// --- Siemens Structured Format ---
DATA_BLOCK "model__HS32_IW50_"
{ S7_Optimized_Access := 'TRUE' }
VERSION :
NON_RETAIN
   VAR
      W_i : ARRAY[0..31, 0..39] OF REAL;
      W_f : ARRAY[0..31, 0..39] OF REAL;
      W_g : ARRAY[0..31, 0..39] OF REAL;
      W_o : ARRAY[0..31, 0..39] OF REAL;
      R_i : ARRAY[0..31, 0..31] OF REAL;
      R_f : ARRAY[0..31, 0..31] OF REAL;
      R_g : ARRAY[0..31, 0..31] OF REAL;
      R_o : ARRAY[0..31, 0..31] OF REAL;
      B_i : ARRAY[0..31] OF REAL;
      B_f : ARRAY[0..31] OF REAL;
      B_g : ARRAY[0..31] OF REAL;
      B_o : ARRAY[0..31] OF REAL;
      FC_W : ARRAY[0..39, 0..31] OF REAL;
      FC_B : ARRAY[0..39] OF REAL;
   END_VAR
BEGIN

      W_i[0,0] := 0.03335211;
      W_i[0,1] := 0.01294965;
      W_i[0,2] := -0.02368959;
      W_i[0,3] := 0.02531582;
      W_i[0,4] := -0.09620859;
      W_i[0,5] := -0.01378066;
      W_i[0,6] := 0.03223424;
      W_i[0,7] := 0.44872370;
      W_i[0,8] := 0.10217454;
      W_i[0,9] := -0.36218736;
      W_i[0,10] := 0.04811719;
      W_i[0,11] := -0.30795375;
      W_i[0,12] := -0.13306537;
      W_i[0,13] := -0.13929474;
      W_i[0,14] := -0.02903975;
      W_i[0,15] := 0.11072005;
      W_i[0,16] := 0.03733860;
      W_i[0,17] := 0.00262149;
      W_i[0,18] := 0.23541802;
      W_i[0,19] := 0.20732951;
      W_i[0,20] := 0.04801108;
      W_i[0,21] := -0.28304836;
      W_i[0,22] := -0.50957590;
      W_i[0,23] := 0.04589643;
      W_i[0,24] := -0.43349111;
      W_i[0,25] := -0.42231610;
      W_i[0,26] := 0.15247093;
      W_i[0,27] := 0.29900289;
      W_i[0,28] := 0.08071815;
      W_i[0,29] := 0.16624704;
      W_i[0,30] := -0.21118966;
      W_i[0,31] := -0.06602232;
      W_i[0,32] := 0.02604864;
      W_i[0,33] := -0.14019786;
      W_i[0,34] := -0.40027091;
      W_i[0,35] := 0.18787135;
      W_i[0,36] := 0.02354476;
      W_i[0,37] := 0.16503902;
      W_i[0,38] := -0.08474749;
      W_i[0,39] := 0.36904612;
      W_i[1,0] := -0.04397624;
      W_i[1,1] := 0.12521634;
      W_i[1,2] := 0.00926329;
      W_i[1,3] := 0.07923686;
      W_i[1,4] := -0.48040998;
      W_i[1,5] := 0.11951946;
      W_i[1,6] := -0.05899520;
      W_i[1,7] := 0.08414336;
      W_i[1,8] := -0.05504049;
      W_i[1,9] := -0.01812936;
      W_i[1,10] := -0.07156652;
      W_i[1,11] := -0.13873386;
      W_i[1,12] := -0.06473546;
      W_i[1,13] := -0.01150122;
      W_i[1,14] := 0.01369441;
      W_i[1,15] := -0.04945480;
      W_i[1,16] := 0.03672740;
      W_i[1,17] := -0.01182620;
      W_i[1,18] := 0.05847014;
      W_i[1,19] := 0.12310074;
      W_i[1,20] := 0.00140591;
      W_i[1,21] := 0.05102165;
      W_i[1,22] := 0.02194597;
      W_i[1,23] := 0.02794340;
      W_i[1,24] := -0.11971385;
      W_i[1,25] := 0.01236170;
      W_i[1,26] := 0.02725715;
      W_i[1,27] := -0.16358410;
      W_i[1,28] := 0.09302291;
      W_i[1,29] := -0.07609808;
      W_i[1,30] := 0.12344577;
      W_i[1,31] := 0.27449563;
      W_i[1,32] := 0.19618334;
      W_i[1,33] := -0.13863903;
      W_i[1,34] := -0.14182809;
      W_i[1,35] := -0.04518571;
      W_i[1,36] := -0.11997688;
      W_i[1,37] := 0.13018343;
      W_i[1,38] := 0.03084990;
      W_i[1,39] := 0.01552542;
      W_i[2,0] := -0.06228839;
      W_i[2,1] := 0.31358635;
      W_i[2,2] := -0.02805484;
      W_i[2,3] := 0.06225382;
      W_i[2,4] := -0.10929245;
      W_i[2,5] := 0.09066710;
      W_i[2,6] := -0.09841387;
      W_i[2,7] := 0.21516874;
      W_i[2,8] := -0.04192384;
      W_i[2,9] := -0.24015123;
      W_i[2,10] := 0.18081841;
      W_i[2,11] := -0.22261326;
      W_i[2,12] := 0.15341285;
      W_i[2,13] := -0.01613901;
      W_i[2,14] := 0.00278526;
      W_i[2,15] := 0.00110682;
      W_i[2,16] := 0.01401542;
      W_i[2,17] := 0.00157240;
      W_i[2,18] := -0.00937896;
      W_i[2,19] := 0.08156285;
      W_i[2,20] := -0.10387972;
      W_i[2,21] := 0.07669238;
      W_i[2,22] := 0.10504947;
      W_i[2,23] := 0.02962043;
      W_i[2,24] := 0.06015503;
      W_i[2,25] := -0.38022354;
      W_i[2,26] := 0.01376416;
      W_i[2,27] := -0.19910932;
      W_i[2,28] := -0.11147632;
      W_i[2,29] := -0.06024737;
      W_i[2,30] := 0.33740976;
      W_i[2,31] := -0.14441007;
      W_i[2,32] := 0.09709183;
      W_i[2,33] := -0.01737254;
      W_i[2,34] := 0.10466792;
      W_i[2,35] := -0.13491732;
      W_i[2,36] := 0.03209321;
      W_i[2,37] := -0.20953350;
      W_i[2,38] := 0.02072377;
      W_i[2,39] := -0.03477554;
      W_i[3,0] := -0.20035338;
      W_i[3,1] := -0.05025988;
      W_i[3,2] := -0.08164182;
      W_i[3,3] := -0.08261910;
      W_i[3,4] := 0.24175876;
      W_i[3,5] := -0.19314556;
      W_i[3,6] := 0.16183864;
      W_i[3,7] := -0.53965092;
      W_i[3,8] := 0.12166216;
      W_i[3,9] := 0.06300285;
      W_i[3,10] := 0.24695574;
      W_i[3,11] := -0.06766498;
      W_i[3,12] := -0.10851647;
      W_i[3,13] := -0.09679550;
      W_i[3,14] := 0.19846407;
      W_i[3,15] := 0.24224226;
      W_i[3,16] := -0.04479418;
      W_i[3,17] := 0.09416196;
      W_i[3,18] := -0.05448310;
      W_i[3,19] := -0.14848493;
      W_i[3,20] := -0.13104467;
      W_i[3,21] := 0.01169914;
      W_i[3,22] := 0.13594244;
      W_i[3,23] := -0.09969987;
      W_i[3,24] := -0.51131010;
      W_i[3,25] := -0.49498364;
      W_i[3,26] := -0.00815858;
      W_i[3,27] := -0.01644909;
      W_i[3,28] := -0.31252897;
      W_i[3,29] := -0.13085435;
      W_i[3,30] := 0.42893934;
      W_i[3,31] := -0.31215337;
      W_i[3,32] := -0.04756459;
      W_i[3,33] := -0.18021715;
      W_i[3,34] := -0.17681709;
      W_i[3,35] := -0.15721944;
      W_i[3,36] := 0.22830988;
      W_i[3,37] := 0.15386219;
      W_i[3,38] := -0.11364616;
      W_i[3,39] := 0.85980165;
      W_i[4,0] := -0.05922852;
      W_i[4,1] := 0.47120315;
      W_i[4,2] := 0.31002536;
      W_i[4,3] := 0.05706808;
      W_i[4,4] := 0.21668130;
      W_i[4,5] := 0.09678623;
      W_i[4,6] := 0.37920210;
      W_i[4,7] := 0.11913582;
      W_i[4,8] := 0.18588071;
      W_i[4,9] := -0.54219109;
      W_i[4,10] := 0.27432936;
      W_i[4,11] := -0.28996110;
      W_i[4,12] := 0.63514346;
      W_i[4,13] := 0.18675460;
      W_i[4,14] := 0.04656186;
      W_i[4,15] := 0.13881819;
      W_i[4,16] := -0.17344026;
      W_i[4,17] := 0.07573078;
      W_i[4,18] := 0.08432268;
      W_i[4,19] := -0.39324254;
      W_i[4,20] := 0.22332989;
      W_i[4,21] := 0.55870950;
      W_i[4,22] := -0.48373845;
      W_i[4,23] := -0.31563666;
      W_i[4,24] := 0.31388757;
      W_i[4,25] := 0.28351381;
      W_i[4,26] := 0.00493392;
      W_i[4,27] := -0.14279558;
      W_i[4,28] := 0.01328408;
      W_i[4,29] := -0.13343237;
      W_i[4,30] := -0.52480948;
      W_i[4,31] := -0.44383386;
      W_i[4,32] := -0.22764747;
      W_i[4,33] := 0.36674559;
      W_i[4,34] := 0.28135881;
      W_i[4,35] := -0.37915036;
      W_i[4,36] := 0.29197508;
      W_i[4,37] := -0.36793157;
      W_i[4,38] := 0.61301214;
      W_i[4,39] := 0.29268816;
      W_i[5,0] := -0.15593423;
      W_i[5,1] := -0.08324785;
      W_i[5,2] := 0.00935801;
      W_i[5,3] := 0.08572404;
      W_i[5,4] := -0.04179911;
      W_i[5,5] := -0.08974203;
      W_i[5,6] := -0.03267067;
      W_i[5,7] := -0.12864745;
      W_i[5,8] := 0.03684423;
      W_i[5,9] := -0.13796446;
      W_i[5,10] := 0.05928193;
      W_i[5,11] := -0.19078448;
      W_i[5,12] := 0.04955722;
      W_i[5,13] := -0.13951716;
      W_i[5,14] := 0.01461054;
      W_i[5,15] := 0.05807864;
      W_i[5,16] := -0.02155071;
      W_i[5,17] := 0.06774671;
      W_i[5,18] := -0.00056143;
      W_i[5,19] := 0.02993268;
      W_i[5,20] := -0.04689442;
      W_i[5,21] := 0.14087728;
      W_i[5,22] := -0.00434205;
      W_i[5,23] := -0.14380206;
      W_i[5,24] := -0.53344935;
      W_i[5,25] := 0.06604308;
      W_i[5,26] := 0.23374112;
      W_i[5,27] := 0.02832700;
      W_i[5,28] := 0.09275237;
      W_i[5,29] := 0.07908134;
      W_i[5,30] := -0.10972932;
      W_i[5,31] := -0.08337840;
      W_i[5,32] := 0.04662216;
      W_i[5,33] := -0.03259875;
      W_i[5,34] := 0.17782964;
      W_i[5,35] := 0.18201338;
      W_i[5,36] := 0.00404544;
      W_i[5,37] := 0.04663613;
      W_i[5,38] := 0.13219389;
      W_i[5,39] := -0.00446346;
      W_i[6,0] := 0.10576568;
      W_i[6,1] := 0.05325136;
      W_i[6,2] := -0.05492130;
      W_i[6,3] := -0.11396622;
      W_i[6,4] := 0.02959487;
      W_i[6,5] := 0.04510606;
      W_i[6,6] := 0.21042347;
      W_i[6,7] := 0.11686674;
      W_i[6,8] := 0.17569162;
      W_i[6,9] := -0.22145574;
      W_i[6,10] := 0.01603481;
      W_i[6,11] := -0.21858092;
      W_i[6,12] := 0.03767690;
      W_i[6,13] := -0.15889299;
      W_i[6,14] := 0.02401877;
      W_i[6,15] := -0.09354293;
      W_i[6,16] := -0.06953581;
      W_i[6,17] := 0.01671052;
      W_i[6,18] := 0.14821531;
      W_i[6,19] := 0.03779463;
      W_i[6,20] := 0.31719235;
      W_i[6,21] := 0.26848948;
      W_i[6,22] := 0.24316274;
      W_i[6,23] := -0.03367342;
      W_i[6,24] := -0.43727583;
      W_i[6,25] := -0.31479907;
      W_i[6,26] := 0.40017867;
      W_i[6,27] := -0.00208360;
      W_i[6,28] := 0.18425919;
      W_i[6,29] := 0.37186173;
      W_i[6,30] := 0.17230935;
      W_i[6,31] := -0.07113405;
      W_i[6,32] := 0.06234986;
      W_i[6,33] := -0.04395010;
      W_i[6,34] := 0.03162268;
      W_i[6,35] := 0.12794030;
      W_i[6,36] := -0.06928633;
      W_i[6,37] := 0.28019226;
      W_i[6,38] := -0.08624983;
      W_i[6,39] := -0.05943641;
      W_i[7,0] := 0.24273345;
      W_i[7,1] := 0.02628726;
      W_i[7,2] := -0.37892520;
      W_i[7,3] := 0.15462431;
      W_i[7,4] := -0.06835640;
      W_i[7,5] := -0.01244921;
      W_i[7,6] := -0.13799721;
      W_i[7,7] := 0.00364937;
      W_i[7,8] := -0.11085126;
      W_i[7,9] := -0.08217847;
      W_i[7,10] := 0.06155964;
      W_i[7,11] := 0.00664949;
      W_i[7,12] := -0.21111001;
      W_i[7,13] := -0.09906641;
      W_i[7,14] := 0.01441233;
      W_i[7,15] := 0.05717637;
      W_i[7,16] := -0.01254125;
      W_i[7,17] := -0.00084031;
      W_i[7,18] := 0.75006574;
      W_i[7,19] := 0.04177287;
      W_i[7,20] := -0.16489621;
      W_i[7,21] := -0.11358984;
      W_i[7,22] := -0.32568359;
      W_i[7,23] := -0.05461695;
      W_i[7,24] := -0.68117988;
      W_i[7,25] := -0.38877121;
      W_i[7,26] := 0.21966200;
      W_i[7,27] := 0.08412468;
      W_i[7,28] := -0.18800470;
      W_i[7,29] := -0.37555104;
      W_i[7,30] := -0.20995075;
      W_i[7,31] := -0.00920301;
      W_i[7,32] := -0.38933340;
      W_i[7,33] := 0.03684454;
      W_i[7,34] := -0.00580212;
      W_i[7,35] := -0.12717755;
      W_i[7,36] := 0.00740355;
      W_i[7,37] := -0.09031770;
      W_i[7,38] := -0.11013316;
      W_i[7,39] := -0.04330545;
      W_i[8,0] := -0.06802954;
      W_i[8,1] := -0.02636882;
      W_i[8,2] := 0.04332832;
      W_i[8,3] := -0.12407507;
      W_i[8,4] := 0.01348176;
      W_i[8,5] := -0.07925858;
      W_i[8,6] := -0.00761013;
      W_i[8,7] := 0.03581184;
      W_i[8,8] := 0.02980794;
      W_i[8,9] := -0.13043974;
      W_i[8,10] := 0.09170759;
      W_i[8,11] := -0.16562377;
      W_i[8,12] := -0.12424939;
      W_i[8,13] := 0.05662967;
      W_i[8,14] := -0.21820237;
      W_i[8,15] := 0.03667807;
      W_i[8,16] := 0.01659469;
      W_i[8,17] := 0.00193780;
      W_i[8,18] := -0.03699196;
      W_i[8,19] := -0.02531029;
      W_i[8,20] := -0.00570031;
      W_i[8,21] := 0.10410964;
      W_i[8,22] := 0.06439263;
      W_i[8,23] := -0.07894669;
      W_i[8,24] := -0.28273982;
      W_i[8,25] := -0.23450002;
      W_i[8,26] := 0.05201263;
      W_i[8,27] := -0.03252214;
      W_i[8,28] := -0.01173223;
      W_i[8,29] := 0.14622457;
      W_i[8,30] := 0.17911775;
      W_i[8,31] := -0.11378439;
      W_i[8,32] := 0.07194026;
      W_i[8,33] := 0.01723621;
      W_i[8,34] := 0.30313444;
      W_i[8,35] := 0.11768141;
      W_i[8,36] := -0.01293503;
      W_i[8,37] := -0.00394995;
      W_i[8,38] := -0.14124557;
      W_i[8,39] := 0.13445212;
      W_i[9,0] := 0.41246179;
      W_i[9,1] := -0.12685674;
      W_i[9,2] := -0.45634085;
      W_i[9,3] := -0.20486909;
      W_i[9,4] := -0.07218436;
      W_i[9,5] := -0.09485383;
      W_i[9,6] := 0.19853495;
      W_i[9,7] := 0.07240235;
      W_i[9,8] := -0.04039089;
      W_i[9,9] := -0.09886632;
      W_i[9,10] := -0.11097286;
      W_i[9,11] := -0.28303620;
      W_i[9,12] := 0.15636595;
      W_i[9,13] := 0.12219298;
      W_i[9,14] := 0.16322424;
      W_i[9,15] := 0.06697550;
      W_i[9,16] := -0.11505034;
      W_i[9,17] := 0.01392226;
      W_i[9,18] := -0.03821991;
      W_i[9,19] := 0.35102692;
      W_i[9,20] := 0.15118374;
      W_i[9,21] := 0.24640937;
      W_i[9,22] := 0.02153728;
      W_i[9,23] := -0.02444457;
      W_i[9,24] := 0.13131861;
      W_i[9,25] := -0.16178758;
      W_i[9,26] := -0.05835283;
      W_i[9,27] := -0.28876659;
      W_i[9,28] := -0.22485775;
      W_i[9,29] := -0.10750232;
      W_i[9,30] := 0.07209923;
      W_i[9,31] := -0.16665789;
      W_i[9,32] := 0.09024238;
      W_i[9,33] := 0.15630057;
      W_i[9,34] := 0.22654596;
      W_i[9,35] := -0.16981296;
      W_i[9,36] := 0.09843912;
      W_i[9,37] := -0.08633557;
      W_i[9,38] := 0.06714951;
      W_i[9,39] := -0.10012744;
      W_i[10,0] := 0.06098233;
      W_i[10,1] := 0.00406449;
      W_i[10,2] := -0.07085112;
      W_i[10,3] := -0.38051835;
      W_i[10,4] := -0.14092854;
      W_i[10,5] := -0.05471934;
      W_i[10,6] := -0.09075350;
      W_i[10,7] := 0.09081808;
      W_i[10,8] := 0.07290499;
      W_i[10,9] := 0.21984702;
      W_i[10,10] := -0.00319992;
      W_i[10,11] := -0.87133026;
      W_i[10,12] := 0.25286415;
      W_i[10,13] := -0.20190343;
      W_i[10,14] := -0.29993787;
      W_i[10,15] := -0.01450086;
      W_i[10,16] := -0.04255661;
      W_i[10,17] := 0.50596321;
      W_i[10,18] := -0.03224555;
      W_i[10,19] := 0.00962685;
      W_i[10,20] := 0.02170906;
      W_i[10,21] := 0.00463841;
      W_i[10,22] := 0.00428250;
      W_i[10,23] := 0.02700867;
      W_i[10,24] := -0.49260652;
      W_i[10,25] := -0.60828519;
      W_i[10,26] := 0.08981935;
      W_i[10,27] := -0.05126838;
      W_i[10,28] := 0.10806957;
      W_i[10,29] := 0.06330517;
      W_i[10,30] := 0.09711373;
      W_i[10,31] := -0.19667481;
      W_i[10,32] := 0.04281054;
      W_i[10,33] := 0.06612559;
      W_i[10,34] := -0.12514877;
      W_i[10,35] := 0.09477433;
      W_i[10,36] := 0.02109047;
      W_i[10,37] := 0.06420635;
      W_i[10,38] := 0.06682578;
      W_i[10,39] := 0.70137119;
      W_i[11,0] := -0.19831482;
      W_i[11,1] := -0.10508762;
      W_i[11,2] := 0.14985219;
      W_i[11,3] := -0.25513422;
      W_i[11,4] := 0.22445941;
      W_i[11,5] := -0.17102213;
      W_i[11,6] := 0.03812301;
      W_i[11,7] := 0.06178447;
      W_i[11,8] := -0.06147041;
      W_i[11,9] := 0.01455363;
      W_i[11,10] := 0.21236670;
      W_i[11,11] := -0.06561671;
      W_i[11,12] := -0.23426783;
      W_i[11,13] := 0.09121598;
      W_i[11,14] := -0.11325682;
      W_i[11,15] := 0.14043726;
      W_i[11,16] := -0.03869899;
      W_i[11,17] := 0.07733488;
      W_i[11,18] := -0.00199524;
      W_i[11,19] := 0.05081591;
      W_i[11,20] := -0.45575571;
      W_i[11,21] := -0.48401207;
      W_i[11,22] := -0.20732693;
      W_i[11,23] := -0.15296169;
      W_i[11,24] := -0.30430803;
      W_i[11,25] := -0.48835382;
      W_i[11,26] := -0.19211042;
      W_i[11,27] := 0.21992902;
      W_i[11,28] := -0.36160839;
      W_i[11,29] := -0.36730286;
      W_i[11,30] := -0.27825427;
      W_i[11,31] := 0.49533325;
      W_i[11,32] := 0.01973951;
      W_i[11,33] := 0.13294254;
      W_i[11,34] := -0.31377479;
      W_i[11,35] := 0.01389581;
      W_i[11,36] := -0.10732657;
      W_i[11,37] := -0.10178760;
      W_i[11,38] := -0.04468285;
      W_i[11,39] := 0.88543254;
      W_i[12,0] := -0.07785182;
      W_i[12,1] := -0.02275736;
      W_i[12,2] := -0.01598639;
      W_i[12,3] := -0.28018406;
      W_i[12,4] := 0.04472728;
      W_i[12,5] := -0.07362497;
      W_i[12,6] := 0.10421625;
      W_i[12,7] := 0.29120883;
      W_i[12,8] := 0.07516699;
      W_i[12,9] := -0.19484363;
      W_i[12,10] := 0.04389035;
      W_i[12,11] := 0.07964118;
      W_i[12,12] := 0.04882551;
      W_i[12,13] := -0.09314007;
      W_i[12,14] := -0.00104783;
      W_i[12,15] := 0.12430931;
      W_i[12,16] := -0.00889617;
      W_i[12,17] := -0.00109596;
      W_i[12,18] := 0.93196803;
      W_i[12,19] := 0.07360591;
      W_i[12,20] := -0.04771593;
      W_i[12,21] := 0.00891263;
      W_i[12,22] := -0.22154218;
      W_i[12,23] := -0.00681991;
      W_i[12,24] := -0.28159559;
      W_i[12,25] := -0.33888876;
      W_i[12,26] := 0.11433282;
      W_i[12,27] := -0.10486361;
      W_i[12,28] := -0.09925523;
      W_i[12,29] := -0.00571722;
      W_i[12,30] := -0.36633971;
      W_i[12,31] := -0.06006427;
      W_i[12,32] := -0.22424956;
      W_i[12,33] := -0.32570857;
      W_i[12,34] := -0.57398140;
      W_i[12,35] := 0.05099113;
      W_i[12,36] := 0.00469301;
      W_i[12,37] := 0.02404906;
      W_i[12,38] := 0.01321469;
      W_i[12,39] := -0.01789427;
      W_i[13,0] := 0.13228506;
      W_i[13,1] := 0.10746437;
      W_i[13,2] := -0.02473475;
      W_i[13,3] := -0.01283106;
      W_i[13,4] := -0.11313344;
      W_i[13,5] := 0.01196120;
      W_i[13,6] := -0.10874924;
      W_i[13,7] := -0.09509301;
      W_i[13,8] := 0.00865637;
      W_i[13,9] := -0.15097018;
      W_i[13,10] := 0.07857790;
      W_i[13,11] := -0.13828419;
      W_i[13,12] := 0.18908830;
      W_i[13,13] := -0.03993330;
      W_i[13,14] := 0.01041046;
      W_i[13,15] := 0.00195818;
      W_i[13,16] := -0.02810182;
      W_i[13,17] := -0.00908193;
      W_i[13,18] := -0.01383985;
      W_i[13,19] := 0.01692491;
      W_i[13,20] := 0.26870248;
      W_i[13,21] := 0.50765073;
      W_i[13,22] := 0.34594440;
      W_i[13,23] := -0.03796029;
      W_i[13,24] := -0.65532976;
      W_i[13,25] := -0.80482006;
      W_i[13,26] := 0.01045384;
      W_i[13,27] := -0.46558616;
      W_i[13,28] := 0.19693999;
      W_i[13,29] := 0.14626113;
      W_i[13,30] := 0.43212712;
      W_i[13,31] := 0.01994485;
      W_i[13,32] := -0.32835758;
      W_i[13,33] := -0.17723863;
      W_i[13,34] := 0.20528001;
      W_i[13,35] := -0.34655216;
      W_i[13,36] := -0.06347063;
      W_i[13,37] := -0.07853378;
      W_i[13,38] := 0.15984800;
      W_i[13,39] := 0.00452000;
      W_i[14,0] := -0.00785071;
      W_i[14,1] := -0.08457682;
      W_i[14,2] := -0.03021882;
      W_i[14,3] := 0.06919254;
      W_i[14,4] := -0.07102513;
      W_i[14,5] := -0.11649032;
      W_i[14,6] := -0.13716960;
      W_i[14,7] := 0.12219854;
      W_i[14,8] := -0.03531046;
      W_i[14,9] := -0.07139499;
      W_i[14,10] := -0.28596520;
      W_i[14,11] := -0.20866406;
      W_i[14,12] := -0.09834762;
      W_i[14,13] := -0.17434466;
      W_i[14,14] := 0.05277216;
      W_i[14,15] := 0.05034710;
      W_i[14,16] := -0.04395842;
      W_i[14,17] := 0.01994520;
      W_i[14,18] := -0.00284745;
      W_i[14,19] := -0.01580888;
      W_i[14,20] := 0.35238999;
      W_i[14,21] := -0.30224216;
      W_i[14,22] := -0.01767650;
      W_i[14,23] := 0.06807997;
      W_i[14,24] := -0.02559922;
      W_i[14,25] := -0.02666317;
      W_i[14,26] := 0.03206453;
      W_i[14,27] := 0.41885376;
      W_i[14,28] := 0.04192250;
      W_i[14,29] := -0.05693231;
      W_i[14,30] := 0.07898923;
      W_i[14,31] := 0.18591896;
      W_i[14,32] := -0.06221836;
      W_i[14,33] := 0.24379699;
      W_i[14,34] := -0.13005574;
      W_i[14,35] := 0.04800267;
      W_i[14,36] := 0.09943730;
      W_i[14,37] := -0.03374345;
      W_i[14,38] := -0.03513518;
      W_i[14,39] := -0.07157569;
      W_i[15,0] := -0.15272453;
      W_i[15,1] := 0.13645852;
      W_i[15,2] := 0.04745365;
      W_i[15,3] := -0.20139949;
      W_i[15,4] := 0.03436549;
      W_i[15,5] := 0.06549827;
      W_i[15,6] := -0.17606948;
      W_i[15,7] := 0.05636362;
      W_i[15,8] := 0.15209863;
      W_i[15,9] := -0.04455522;
      W_i[15,10] := 0.01616382;
      W_i[15,11] := 0.02472791;
      W_i[15,12] := 0.01587282;
      W_i[15,13] := 0.06205805;
      W_i[15,14] := -0.01110538;
      W_i[15,15] := -0.05222612;
      W_i[15,16] := -0.00958592;
      W_i[15,17] := 0.05923622;
      W_i[15,18] := 0.03878036;
      W_i[15,19] := -0.04121817;
      W_i[15,20] := -0.04009682;
      W_i[15,21] := 0.02127116;
      W_i[15,22] := -0.04295387;
      W_i[15,23] := -0.08172908;
      W_i[15,24] := -0.48291191;
      W_i[15,25] := -0.58466184;
      W_i[15,26] := -0.04407280;
      W_i[15,27] := 0.00633614;
      W_i[15,28] := -0.10225561;
      W_i[15,29] := 0.48959246;
      W_i[15,30] := -0.22612220;
      W_i[15,31] := -0.01089828;
      W_i[15,32] := -0.25822705;
      W_i[15,33] := -0.17706192;
      W_i[15,34] := -0.61160076;
      W_i[15,35] := 0.09040477;
      W_i[15,36] := 0.02512925;
      W_i[15,37] := -0.06701392;
      W_i[15,38] := -0.08561996;
      W_i[15,39] := 0.53837699;
      W_i[16,0] := -0.07811758;
      W_i[16,1] := 0.05202470;
      W_i[16,2] := 0.03025672;
      W_i[16,3] := 0.04235693;
      W_i[16,4] := -0.06725603;
      W_i[16,5] := -0.00081394;
      W_i[16,6] := -0.09191743;
      W_i[16,7] := 0.24823768;
      W_i[16,8] := 0.02800119;
      W_i[16,9] := -0.27142274;
      W_i[16,10] := -0.06025495;
      W_i[16,11] := -0.51023978;
      W_i[16,12] := 0.54432988;
      W_i[16,13] := -0.07693134;
      W_i[16,14] := 0.03643584;
      W_i[16,15] := 0.04252481;
      W_i[16,16] := -0.00319035;
      W_i[16,17] := -0.16166179;
      W_i[16,18] := -0.10264453;
      W_i[16,19] := -0.72658694;
      W_i[16,20] := -0.08637008;
      W_i[16,21] := -0.15963581;
      W_i[16,22] := -0.16920443;
      W_i[16,23] := -0.03855850;
      W_i[16,24] := -0.09449768;
      W_i[16,25] := -0.15130939;
      W_i[16,26] := -0.07037468;
      W_i[16,27] := 0.05760185;
      W_i[16,28] := 0.01705931;
      W_i[16,29] := 0.05011314;
      W_i[16,30] := -0.01099099;
      W_i[16,31] := -0.06498095;
      W_i[16,32] := 0.15388052;
      W_i[16,33] := -0.03008743;
      W_i[16,34] := -0.91294670;
      W_i[16,35] := 0.04827264;
      W_i[16,36] := 0.00881240;
      W_i[16,37] := 0.02179604;
      W_i[16,38] := 0.47361013;
      W_i[16,39] := 0.58336878;
      W_i[17,0] := -0.22612889;
      W_i[17,1] := -0.03230098;
      W_i[17,2] := 0.24163076;
      W_i[17,3] := 0.20527579;
      W_i[17,4] := -0.44036463;
      W_i[17,5] := 0.28084049;
      W_i[17,6] := -0.51067066;
      W_i[17,7] := 0.07827551;
      W_i[17,8] := -0.09376909;
      W_i[17,9] := -0.11010143;
      W_i[17,10] := -0.31384867;
      W_i[17,11] := -0.58446574;
      W_i[17,12] := -0.01893969;
      W_i[17,13] := -0.05360400;
      W_i[17,14] := 0.07922329;
      W_i[17,15] := -0.01531055;
      W_i[17,16] := 0.16111493;
      W_i[17,17] := 0.20549683;
      W_i[17,18] := 0.35656574;
      W_i[17,19] := 0.11651949;
      W_i[17,20] := 0.09743474;
      W_i[17,21] := 0.14924602;
      W_i[17,22] := 0.13436577;
      W_i[17,23] := 0.04628479;
      W_i[17,24] := -0.27565825;
      W_i[17,25] := -0.53178447;
      W_i[17,26] := -0.07750764;
      W_i[17,27] := -0.00472372;
      W_i[17,28] := 0.36722642;
      W_i[17,29] := -0.59928131;
      W_i[17,30] := 0.19017772;
      W_i[17,31] := -0.13342376;
      W_i[17,32] := 0.06940365;
      W_i[17,33] := 0.19215287;
      W_i[17,34] := -0.27029362;
      W_i[17,35] := 0.32601219;
      W_i[17,36] := 0.06043479;
      W_i[17,37] := 0.03219402;
      W_i[17,38] := -0.06975342;
      W_i[17,39] := 0.23071089;
      W_i[18,0] := 0.40103209;
      W_i[18,1] := 0.04176520;
      W_i[18,2] := -0.13692427;
      W_i[18,3] := -0.07025969;
      W_i[18,4] := 0.18873395;
      W_i[18,5] := -0.04070675;
      W_i[18,6] := -0.20584334;
      W_i[18,7] := -0.01120962;
      W_i[18,8] := -0.19570278;
      W_i[18,9] := 0.29601005;
      W_i[18,10] := -0.11879414;
      W_i[18,11] := 0.17400281;
      W_i[18,12] := 0.00161714;
      W_i[18,13] := -0.08103235;
      W_i[18,14] := 0.21251068;
      W_i[18,15] := 0.01489939;
      W_i[18,16] := 0.04055646;
      W_i[18,17] := 0.04331359;
      W_i[18,18] := 0.00444761;
      W_i[18,19] := -0.62320471;
      W_i[18,20] := -0.16792732;
      W_i[18,21] := 0.13485593;
      W_i[18,22] := -0.09223303;
      W_i[18,23] := 0.01478722;
      W_i[18,24] := -0.68178695;
      W_i[18,25] := -0.42708310;
      W_i[18,26] := 0.45379946;
      W_i[18,27] := 0.20425461;
      W_i[18,28] := -0.21162227;
      W_i[18,29] := 0.10539333;
      W_i[18,30] := -0.09736414;
      W_i[18,31] := -0.51747489;
      W_i[18,32] := 0.09172474;
      W_i[18,33] := 0.19873166;
      W_i[18,34] := -0.02417281;
      W_i[18,35] := 0.23588333;
      W_i[18,36] := -0.14076033;
      W_i[18,37] := 0.46431357;
      W_i[18,38] := 0.09138855;
      W_i[18,39] := 0.86890060;
      W_i[19,0] := -0.06011394;
      W_i[19,1] := -0.01500004;
      W_i[19,2] := -0.04331917;
      W_i[19,3] := 0.18670803;
      W_i[19,4] := 0.12613097;
      W_i[19,5] := 0.00880916;
      W_i[19,6] := -0.02774461;
      W_i[19,7] := -0.14737256;
      W_i[19,8] := 0.03255391;
      W_i[19,9] := 0.01357013;
      W_i[19,10] := 0.02901205;
      W_i[19,11] := -0.09940059;
      W_i[19,12] := -0.17535669;
      W_i[19,13] := -0.16476427;
      W_i[19,14] := -0.03231515;
      W_i[19,15] := 0.29976013;
      W_i[19,16] := -0.22633493;
      W_i[19,17] := 0.04706604;
      W_i[19,18] := -0.04980571;
      W_i[19,19] := 0.04330605;
      W_i[19,20] := -0.06072775;
      W_i[19,21] := -0.15681855;
      W_i[19,22] := -0.17704034;
      W_i[19,23] := -0.00916669;
      W_i[19,24] := 0.10120902;
      W_i[19,25] := -0.01640362;
      W_i[19,26] := 0.07318049;
      W_i[19,27] := 0.21290408;
      W_i[19,28] := -0.27156901;
      W_i[19,29] := -0.02253475;
      W_i[19,30] := -0.28479761;
      W_i[19,31] := 0.05325111;
      W_i[19,32] := -0.05720755;
      W_i[19,33] := -0.06733356;
      W_i[19,34] := -0.48600927;
      W_i[19,35] := -0.02064243;
      W_i[19,36] := -0.06231465;
      W_i[19,37] := 0.11734369;
      W_i[19,38] := 0.30606124;
      W_i[19,39] := 0.75707734;
      W_i[20,0] := -0.21834370;
      W_i[20,1] := -0.37634116;
      W_i[20,2] := 0.37927234;
      W_i[20,3] := 0.18053402;
      W_i[20,4] := -0.11320233;
      W_i[20,5] := -0.11718341;
      W_i[20,6] := 0.05376241;
      W_i[20,7] := 0.02935014;
      W_i[20,8] := 0.00259118;
      W_i[20,9] := -0.16540758;
      W_i[20,10] := 0.07926913;
      W_i[20,11] := -0.30344686;
      W_i[20,12] := -0.15024255;
      W_i[20,13] := 0.12091222;
      W_i[20,14] := 0.03411222;
      W_i[20,15] := -0.05019326;
      W_i[20,16] := 0.02392713;
      W_i[20,17] := -0.02823546;
      W_i[20,18] := 0.00852875;
      W_i[20,19] := 0.05116982;
      W_i[20,20] := -0.07963332;
      W_i[20,21] := 0.25724292;
      W_i[20,22] := -0.09602219;
      W_i[20,23] := -0.08398317;
      W_i[20,24] := 0.23696989;
      W_i[20,25] := 0.25781205;
      W_i[20,26] := -0.04276172;
      W_i[20,27] := -0.56399757;
      W_i[20,28] := -0.03985150;
      W_i[20,29] := 0.08735032;
      W_i[20,30] := 0.11606380;
      W_i[20,31] := 0.10737984;
      W_i[20,32] := -0.05359823;
      W_i[20,33] := 0.02176436;
      W_i[20,34] := 0.10568735;
      W_i[20,35] := 0.15294984;
      W_i[20,36] := -0.07409501;
      W_i[20,37] := -0.01986608;
      W_i[20,38] := 0.10280561;
      W_i[20,39] := 0.00202793;
      W_i[21,0] := 0.01244066;
      W_i[21,1] := -0.08776394;
      W_i[21,2] := 0.00320476;
      W_i[21,3] := -0.04366220;
      W_i[21,4] := -0.04889725;
      W_i[21,5] := -0.03951695;
      W_i[21,6] := 0.06806803;
      W_i[21,7] := -0.15357529;
      W_i[21,8] := 0.00562375;
      W_i[21,9] := -0.08162130;
      W_i[21,10] := 0.00548499;
      W_i[21,11] := -0.09151895;
      W_i[21,12] := -0.00889677;
      W_i[21,13] := -0.12972501;
      W_i[21,14] := -0.00167885;
      W_i[21,15] := -0.00695266;
      W_i[21,16] := 0.01370465;
      W_i[21,17] := -0.00067664;
      W_i[21,18] := 0.05669603;
      W_i[21,19] := 0.00472060;
      W_i[21,20] := -0.09169029;
      W_i[21,21] := -0.13030174;
      W_i[21,22] := 0.11552692;
      W_i[21,23] := -0.12622538;
      W_i[21,24] := -0.45613086;
      W_i[21,25] := -0.30946380;
      W_i[21,26] := 0.12234695;
      W_i[21,27] := -0.01556969;
      W_i[21,28] := -0.06982312;
      W_i[21,29] := 0.19435593;
      W_i[21,30] := -0.08212201;
      W_i[21,31] := -0.08049136;
      W_i[21,32] := -0.05780566;
      W_i[21,33] := 0.04121880;
      W_i[21,34] := -0.52323383;
      W_i[21,35] := 0.25505278;
      W_i[21,36] := -0.01052439;
      W_i[21,37] := 0.19438845;
      W_i[21,38] := 0.00495974;
      W_i[21,39] := 0.01865052;
      W_i[22,0] := 0.13598847;
      W_i[22,1] := -0.00137104;
      W_i[22,2] := -0.14428510;
      W_i[22,3] := -0.08302084;
      W_i[22,4] := -0.20576182;
      W_i[22,5] := -0.01815082;
      W_i[22,6] := -0.13738698;
      W_i[22,7] := -0.09441074;
      W_i[22,8] := 0.12739091;
      W_i[22,9] := -0.15741669;
      W_i[22,10] := 0.05683972;
      W_i[22,11] := -0.23765637;
      W_i[22,12] := 0.02600284;
      W_i[22,13] := -0.20088109;
      W_i[22,14] := 0.09838137;
      W_i[22,15] := -0.25285217;
      W_i[22,16] := -0.02274646;
      W_i[22,17] := -0.04241041;
      W_i[22,18] := 0.06986310;
      W_i[22,19] := 0.01868251;
      W_i[22,20] := 0.12563545;
      W_i[22,21] := 0.05377704;
      W_i[22,22] := 0.18017660;
      W_i[22,23] := 0.04133203;
      W_i[22,24] := 0.34861264;
      W_i[22,25] := 0.53120559;
      W_i[22,26] := 0.10605080;
      W_i[22,27] := 0.01764100;
      W_i[22,28] := -0.17181937;
      W_i[22,29] := -0.22923233;
      W_i[22,30] := -0.07923669;
      W_i[22,31] := -0.05656500;
      W_i[22,32] := 0.13083638;
      W_i[22,33] := 0.04422931;
      W_i[22,34] := 0.03540160;
      W_i[22,35] := -0.08169101;
      W_i[22,36] := 0.01437967;
      W_i[22,37] := 0.01002266;
      W_i[22,38] := 0.17844988;
      W_i[22,39] := 0.44851547;
      W_i[23,0] := -0.11353187;
      W_i[23,1] := 0.13802458;
      W_i[23,2] := 0.04801157;
      W_i[23,3] := 0.19126737;
      W_i[23,4] := -0.02774257;
      W_i[23,5] := -0.11002547;
      W_i[23,6] := -0.07597420;
      W_i[23,7] := 0.07305055;
      W_i[23,8] := -0.02948767;
      W_i[23,9] := 0.06787046;
      W_i[23,10] := -0.13287917;
      W_i[23,11] := -0.23878390;
      W_i[23,12] := -0.16946453;
      W_i[23,13] := -0.01882853;
      W_i[23,14] := 0.00419446;
      W_i[23,15] := -0.02854069;
      W_i[23,16] := 0.03501445;
      W_i[23,17] := -0.02042479;
      W_i[23,18] := 0.03517327;
      W_i[23,19] := 0.06832731;
      W_i[23,20] := 0.08877181;
      W_i[23,21] := -0.13232544;
      W_i[23,22] := 0.03553335;
      W_i[23,23] := -0.17476059;
      W_i[23,24] := -0.13496134;
      W_i[23,25] := 0.06990138;
      W_i[23,26] := 0.03886210;
      W_i[23,27] := -0.10751740;
      W_i[23,28] := -0.00182543;
      W_i[23,29] := 0.06371216;
      W_i[23,30] := 0.00089110;
      W_i[23,31] := 0.29507750;
      W_i[23,32] := 0.16118304;
      W_i[23,33] := 0.05159265;
      W_i[23,34] := 0.02121187;
      W_i[23,35] := -0.11368499;
      W_i[23,36] := 0.09601352;
      W_i[23,37] := -0.03368830;
      W_i[23,38] := -0.09560180;
      W_i[23,39] := 0.04410608;
      W_i[24,0] := 0.12907231;
      W_i[24,1] := 0.00349400;
      W_i[24,2] := -0.03250685;
      W_i[24,3] := -0.11876480;
      W_i[24,4] := -0.09973786;
      W_i[24,5] := 0.12441619;
      W_i[24,6] := 0.18852201;
      W_i[24,7] := 0.08817047;
      W_i[24,8] := 0.05041340;
      W_i[24,9] := -0.16866046;
      W_i[24,10] := 0.05290342;
      W_i[24,11] := -0.14306267;
      W_i[24,12] := 0.07523957;
      W_i[24,13] := -0.03941730;
      W_i[24,14] := 0.00118544;
      W_i[24,15] := -0.05347997;
      W_i[24,16] := -0.01991534;
      W_i[24,17] := 0.01214673;
      W_i[24,18] := 0.05419031;
      W_i[24,19] := 0.05075099;
      W_i[24,20] := 0.28088364;
      W_i[24,21] := 0.21089576;
      W_i[24,22] := 0.05161647;
      W_i[24,23] := -0.12937893;
      W_i[24,24] := -0.88216209;
      W_i[24,25] := -0.45865399;
      W_i[24,26] := 0.13305612;
      W_i[24,27] := -0.26171306;
      W_i[24,28] := 0.02579498;
      W_i[24,29] := 0.06367037;
      W_i[24,30] := 0.06579091;
      W_i[24,31] := -0.05059954;
      W_i[24,32] := -0.03575664;
      W_i[24,33] := -0.23555161;
      W_i[24,34] := 0.14354263;
      W_i[24,35] := 0.04409879;
      W_i[24,36] := -0.05239694;
      W_i[24,37] := 0.14840053;
      W_i[24,38] := 0.01412896;
      W_i[24,39] := 0.03093194;
      W_i[25,0] := -0.10782371;
      W_i[25,1] := -0.01355948;
      W_i[25,2] := 0.07241292;
      W_i[25,3] := -0.16890974;
      W_i[25,4] := 0.11865858;
      W_i[25,5] := 0.09844998;
      W_i[25,6] := 0.25812393;
      W_i[25,7] := -0.17237015;
      W_i[25,8] := -0.20769525;
      W_i[25,9] := 0.08842477;
      W_i[25,10] := 0.12996043;
      W_i[25,11] := -0.79491919;
      W_i[25,12] := 0.74928349;
      W_i[25,13] := -0.05475974;
      W_i[25,14] := -0.00581676;
      W_i[25,15] := -1.19459748;
      W_i[25,16] := -0.06734265;
      W_i[25,17] := 0.31761691;
      W_i[25,18] := 0.26755145;
      W_i[25,19] := 0.43190241;
      W_i[25,20] := 0.07431526;
      W_i[25,21] := 0.63314551;
      W_i[25,22] := -0.19244106;
      W_i[25,23] := 0.07679500;
      W_i[25,24] := 0.48746341;
      W_i[25,25] := 0.39778945;
      W_i[25,26] := -0.09085509;
      W_i[25,27] := -0.25928289;
      W_i[25,28] := 0.01539844;
      W_i[25,29] := -0.12492942;
      W_i[25,30] := 0.05111655;
      W_i[25,31] := 0.14279488;
      W_i[25,32] := -0.00017076;
      W_i[25,33] := 0.08198984;
      W_i[25,34] := -0.25336066;
      W_i[25,35] := 0.09243240;
      W_i[25,36] := -0.09799714;
      W_i[25,37] := -0.22570664;
      W_i[25,38] := 0.07282528;
      W_i[25,39] := -0.17275944;
      W_i[26,0] := 0.14802153;
      W_i[26,1] := 0.49659914;
      W_i[26,2] := -0.22974068;
      W_i[26,3] := -0.11983906;
      W_i[26,4] := 0.13968794;
      W_i[26,5] := 0.29743901;
      W_i[26,6] := 0.33969167;
      W_i[26,7] := 0.19421862;
      W_i[26,8] := -0.30833629;
      W_i[26,9] := 0.28232381;
      W_i[26,10] := -0.64658439;
      W_i[26,11] := -0.16491407;
      W_i[26,12] := -0.32558659;
      W_i[26,13] := 0.72759610;
      W_i[26,14] := 0.27591926;
      W_i[26,15] := -0.37322342;
      W_i[26,16] := 0.05170191;
      W_i[26,17] := -0.39006528;
      W_i[26,18] := 1.02482784;
      W_i[26,19] := -0.36565745;
      W_i[26,20] := -0.44499063;
      W_i[26,21] := 0.06149385;
      W_i[26,22] := 0.00500516;
      W_i[26,23] := 1.19761324;
      W_i[26,24] := -0.02737883;
      W_i[26,25] := 0.13198939;
      W_i[26,26] := -0.01217330;
      W_i[26,27] := 0.52076274;
      W_i[26,28] := -0.41753161;
      W_i[26,29] := -0.08724838;
      W_i[26,30] := -0.02137602;
      W_i[26,31] := -0.10584451;
      W_i[26,32] := -0.15371148;
      W_i[26,33] := -0.13383582;
      W_i[26,34] := -0.14327239;
      W_i[26,35] := -0.01230759;
      W_i[26,36] := 0.04848051;
      W_i[26,37] := -0.07385743;
      W_i[26,38] := 0.39123389;
      W_i[26,39] := -0.20425555;
      W_i[27,0] := 0.14738478;
      W_i[27,1] := 0.05069282;
      W_i[27,2] := -0.13511746;
      W_i[27,3] := -0.18692465;
      W_i[27,4] := -0.02400398;
      W_i[27,5] := -0.08836709;
      W_i[27,6] := 0.14841202;
      W_i[27,7] := 0.36201897;
      W_i[27,8] := 0.13706896;
      W_i[27,9] := -0.18912838;
      W_i[27,10] := -0.06113405;
      W_i[27,11] := -0.08270318;
      W_i[27,12] := -0.03695736;
      W_i[27,13] := -0.02962635;
      W_i[27,14] := 0.00381610;
      W_i[27,15] := 0.00979117;
      W_i[27,16] := 0.13083130;
      W_i[27,17] := -0.10384305;
      W_i[27,18] := 0.00907254;
      W_i[27,19] := 0.13926661;
      W_i[27,20] := 0.14822160;
      W_i[27,21] := 0.21821545;
      W_i[27,22] := 0.01221289;
      W_i[27,23] := 0.00253812;
      W_i[27,24] := -0.40003973;
      W_i[27,25] := 0.03202270;
      W_i[27,26] := 0.03787104;
      W_i[27,27] := -0.20770845;
      W_i[27,28] := 0.06803070;
      W_i[27,29] := 0.03431870;
      W_i[27,30] := 0.12083164;
      W_i[27,31] := -0.04855001;
      W_i[27,32] := 0.03430030;
      W_i[27,33] := -0.16165301;
      W_i[27,34] := 0.18641113;
      W_i[27,35] := 0.06492400;
      W_i[27,36] := 0.00585721;
      W_i[27,37] := 0.04836555;
      W_i[27,38] := -0.00242327;
      W_i[27,39] := -0.00128781;
      W_i[28,0] := -0.08962595;
      W_i[28,1] := -0.07614843;
      W_i[28,2] := 0.10791972;
      W_i[28,3] := -0.13034192;
      W_i[28,4] := -0.04829107;
      W_i[28,5] := -0.16795525;
      W_i[28,6] := 0.03756035;
      W_i[28,7] := -0.35099345;
      W_i[28,8] := 0.00150952;
      W_i[28,9] := 0.28438553;
      W_i[28,10] := -0.11453783;
      W_i[28,11] := -0.16691865;
      W_i[28,12] := -0.06418688;
      W_i[28,13] := -0.23560973;
      W_i[28,14] := 0.03788418;
      W_i[28,15] := -0.02843215;
      W_i[28,16] := -0.15510513;
      W_i[28,17] := -0.02401991;
      W_i[28,18] := 0.10050558;
      W_i[28,19] := -0.08189131;
      W_i[28,20] := -0.04796758;
      W_i[28,21] := 0.14852434;
      W_i[28,22] := 0.17933218;
      W_i[28,23] := 0.03969023;
      W_i[28,24] := 0.12722230;
      W_i[28,25] := 0.18355598;
      W_i[28,26] := 0.04152403;
      W_i[28,27] := -0.00643694;
      W_i[28,28] := 0.08877222;
      W_i[28,29] := 0.22853936;
      W_i[28,30] := -0.05319020;
      W_i[28,31] := 0.03955037;
      W_i[28,32] := 0.05882454;
      W_i[28,33] := 0.00072954;
      W_i[28,34] := 0.10105743;
      W_i[28,35] := 0.11781047;
      W_i[28,36] := 0.06220448;
      W_i[28,37] := 0.25568888;
      W_i[28,38] := -0.11655334;
      W_i[28,39] := 1.13950896;
      W_i[29,0] := -0.02707428;
      W_i[29,1] := -0.18842031;
      W_i[29,2] := -0.09791464;
      W_i[29,3] := -0.11183339;
      W_i[29,4] := -0.15648490;
      W_i[29,5] := 0.00410932;
      W_i[29,6] := 0.02442070;
      W_i[29,7] := -0.30917168;
      W_i[29,8] := -0.00766938;
      W_i[29,9] := 0.09439659;
      W_i[29,10] := 0.05856450;
      W_i[29,11] := -0.05623395;
      W_i[29,12] := 0.13410486;
      W_i[29,13] := -0.51531732;
      W_i[29,14] := 0.00582052;
      W_i[29,15] := 0.01077591;
      W_i[29,16] := -0.03078771;
      W_i[29,17] := 0.01352735;
      W_i[29,18] := 0.29730627;
      W_i[29,19] := 0.00708061;
      W_i[29,20] := -0.05041182;
      W_i[29,21] := -0.28822875;
      W_i[29,22] := -0.15998779;
      W_i[29,23] := 0.26153132;
      W_i[29,24] := -0.71995407;
      W_i[29,25] := -0.80026358;
      W_i[29,26] := 0.15403639;
      W_i[29,27] := -0.01868674;
      W_i[29,28] := -0.00473319;
      W_i[29,29] := -0.17840651;
      W_i[29,30] := -0.04518585;
      W_i[29,31] := 0.03597238;
      W_i[29,32] := 0.32715401;
      W_i[29,33] := 0.14597069;
      W_i[29,34] := -0.11820438;
      W_i[29,35] := -0.03648159;
      W_i[29,36] := -0.03277907;
      W_i[29,37] := -0.04239029;
      W_i[29,38] := 0.03452786;
      W_i[29,39] := -0.02934660;
      W_i[30,0] := -0.07876550;
      W_i[30,1] := -0.08495881;
      W_i[30,2] := -0.01209893;
      W_i[30,3] := -0.27028769;
      W_i[30,4] := 0.13052113;
      W_i[30,5] := -0.04665546;
      W_i[30,6] := -0.06021402;
      W_i[30,7] := -0.22987078;
      W_i[30,8] := 0.22273731;
      W_i[30,9] := 0.18734318;
      W_i[30,10] := -0.04719684;
      W_i[30,11] := 0.31970531;
      W_i[30,12] := -0.21497457;
      W_i[30,13] := 0.11974692;
      W_i[30,14] := 0.12075783;
      W_i[30,15] := -0.01226926;
      W_i[30,16] := -0.25517735;
      W_i[30,17] := -0.08420363;
      W_i[30,18] := -0.02085932;
      W_i[30,19] := 0.09974496;
      W_i[30,20] := -0.16216479;
      W_i[30,21] := 0.11611823;
      W_i[30,22] := 0.03156393;
      W_i[30,23] := 0.00782066;
      W_i[30,24] := 0.14692961;
      W_i[30,25] := -0.14290850;
      W_i[30,26] := -0.06736486;
      W_i[30,27] := 0.35548598;
      W_i[30,28] := 0.16093346;
      W_i[30,29] := -0.03011825;
      W_i[30,30] := 0.09389694;
      W_i[30,31] := 0.08177742;
      W_i[30,32] := -0.11979201;
      W_i[30,33] := -0.09875193;
      W_i[30,34] := -0.82327485;
      W_i[30,35] := -0.15285930;
      W_i[30,36] := 0.01101867;
      W_i[30,37] := -0.09208991;
      W_i[30,38] := 0.09232371;
      W_i[30,39] := 0.19146815;
      W_i[31,0] := 0.03494624;
      W_i[31,1] := 0.59522063;
      W_i[31,2] := -0.04113444;
      W_i[31,3] := 0.01630584;
      W_i[31,4] := -0.02753457;
      W_i[31,5] := -0.02803145;
      W_i[31,6] := 0.02850694;
      W_i[31,7] := -0.03007192;
      W_i[31,8] := 0.03410652;
      W_i[31,9] := 0.08756022;
      W_i[31,10] := 0.06637421;
      W_i[31,11] := 0.04986396;
      W_i[31,12] := -0.22093016;
      W_i[31,13] := 0.01523994;
      W_i[31,14] := 0.00753404;
      W_i[31,15] := 0.03791665;
      W_i[31,16] := 0.00949601;
      W_i[31,17] := 0.01877867;
      W_i[31,18] := -0.00670868;
      W_i[31,19] := 0.02808223;
      W_i[31,20] := 0.16238739;
      W_i[31,21] := 0.22188728;
      W_i[31,22] := 0.05416815;
      W_i[31,23] := -0.08576757;
      W_i[31,24] := -0.06725195;
      W_i[31,25] := 0.16834541;
      W_i[31,26] := 0.00612936;
      W_i[31,27] := -0.08754817;
      W_i[31,28] := -0.12403286;
      W_i[31,29] := 0.12124602;
      W_i[31,30] := 0.11540975;
      W_i[31,31] := 0.20918615;
      W_i[31,32] := -0.05494162;
      W_i[31,33] := 0.15834704;
      W_i[31,34] := -0.02028835;
      W_i[31,35] := 0.05372176;
      W_i[31,36] := 0.00309684;
      W_i[31,37] := -0.07195709;
      W_i[31,38] := 0.01512725;
      W_i[31,39] := -0.01948231;
      W_f[0,0] := 0.51486415;
      W_f[0,1] := 0.08947392;
      W_f[0,2] := -0.36361036;
      W_f[0,3] := 0.09339785;
      W_f[0,4] := 0.14571777;
      W_f[0,5] := 0.06567094;
      W_f[0,6] := 0.00099035;
      W_f[0,7] := 0.11427882;
      W_f[0,8] := 0.00807121;
      W_f[0,9] := 0.21890542;
      W_f[0,10] := -0.64552224;
      W_f[0,11] := 0.48954877;
      W_f[0,12] := -0.42364863;
      W_f[0,13] := 0.58121473;
      W_f[0,14] := -0.14598204;
      W_f[0,15] := 0.00128960;
      W_f[0,16] := 0.03425161;
      W_f[0,17] := 1.12171865;
      W_f[0,18] := 1.12738287;
      W_f[0,19] := -0.37528831;
      W_f[0,20] := -0.20803723;
      W_f[0,21] := -0.05376172;
      W_f[0,22] := -0.18022813;
      W_f[0,23] := -0.02734460;
      W_f[0,24] := 0.48543248;
      W_f[0,25] := 0.75121063;
      W_f[0,26] := -0.30286953;
      W_f[0,27] := 0.31402928;
      W_f[0,28] := -0.10319208;
      W_f[0,29] := -0.00672843;
      W_f[0,30] := -0.10800045;
      W_f[0,31] := -0.10890652;
      W_f[0,32] := 0.00558155;
      W_f[0,33] := 0.05390153;
      W_f[0,34] := 0.21246098;
      W_f[0,35] := -0.13201155;
      W_f[0,36] := 0.13524032;
      W_f[0,37] := -0.07276954;
      W_f[0,38] := -0.19470990;
      W_f[0,39] := -0.11452613;
      W_f[1,0] := -0.05178328;
      W_f[1,1] := -0.06958245;
      W_f[1,2] := -0.00605204;
      W_f[1,3] := 0.36955360;
      W_f[1,4] := 0.17416821;
      W_f[1,5] := -0.31491226;
      W_f[1,6] := -0.18974228;
      W_f[1,7] := -0.29025239;
      W_f[1,8] := 0.03730386;
      W_f[1,9] := -0.38043457;
      W_f[1,10] := -0.01308284;
      W_f[1,11] := 0.22701837;
      W_f[1,12] := 0.20134453;
      W_f[1,13] := 0.16289818;
      W_f[1,14] := 0.00762439;
      W_f[1,15] := -0.23973660;
      W_f[1,16] := -0.00415309;
      W_f[1,17] := 0.02410719;
      W_f[1,18] := -0.15452637;
      W_f[1,19] := -0.16436656;
      W_f[1,20] := -0.63187164;
      W_f[1,21] := -0.28277576;
      W_f[1,22] := -0.04835546;
      W_f[1,23] := -0.08373724;
      W_f[1,24] := -0.21453397;
      W_f[1,25] := -0.21943620;
      W_f[1,26] := -0.33646676;
      W_f[1,27] := 0.36604458;
      W_f[1,28] := -0.13385138;
      W_f[1,29] := -0.16978027;
      W_f[1,30] := -0.04827464;
      W_f[1,31] := -0.12681709;
      W_f[1,32] := -0.01190789;
      W_f[1,33] := -0.09755614;
      W_f[1,34] := -0.00193382;
      W_f[1,35] := -0.10313755;
      W_f[1,36] := -0.18212183;
      W_f[1,37] := 0.03042977;
      W_f[1,38] := -0.05414731;
      W_f[1,39] := 0.23028247;
      W_f[2,0] := -0.21537660;
      W_f[2,1] := 0.64421695;
      W_f[2,2] := 0.11080614;
      W_f[2,3] := -0.02968636;
      W_f[2,4] := -0.14276281;
      W_f[2,5] := 0.10779046;
      W_f[2,6] := -0.23214811;
      W_f[2,7] := -0.21947241;
      W_f[2,8] := -0.24958789;
      W_f[2,9] := 0.06077507;
      W_f[2,10] := -0.04725618;
      W_f[2,11] := -0.15846497;
      W_f[2,12] := -0.40300497;
      W_f[2,13] := -0.21110040;
      W_f[2,14] := -0.07022974;
      W_f[2,15] := -0.23936947;
      W_f[2,16] := -0.13589548;
      W_f[2,17] := 0.44120890;
      W_f[2,18] := -0.01683923;
      W_f[2,19] := -0.19376102;
      W_f[2,20] := -0.12328323;
      W_f[2,21] := 0.21011120;
      W_f[2,22] := 0.07557736;
      W_f[2,23] := 0.19787639;
      W_f[2,24] := 1.72647262;
      W_f[2,25] := 1.69331408;
      W_f[2,26] := -0.17228767;
      W_f[2,27] := 0.30382201;
      W_f[2,28] := 0.11962258;
      W_f[2,29] := 0.00382000;
      W_f[2,30] := -0.08143448;
      W_f[2,31] := -0.30318356;
      W_f[2,32] := 0.02209908;
      W_f[2,33] := -0.01385949;
      W_f[2,34] := 0.43391925;
      W_f[2,35] := -0.26671097;
      W_f[2,36] := -0.17454998;
      W_f[2,37] := -0.29695323;
      W_f[2,38] := 0.23935039;
      W_f[2,39] := 0.05324025;
      W_f[3,0] := -0.88779169;
      W_f[3,1] := 0.16894802;
      W_f[3,2] := 0.27028313;
      W_f[3,3] := -1.06181979;
      W_f[3,4] := 0.26275194;
      W_f[3,5] := -0.51793051;
      W_f[3,6] := 0.76576924;
      W_f[3,7] := 0.35057229;
      W_f[3,8] := 0.47874117;
      W_f[3,9] := 0.21663344;
      W_f[3,10] := 0.75385141;
      W_f[3,11] := -0.31677344;
      W_f[3,12] := -0.12540899;
      W_f[3,13] := -0.11491809;
      W_f[3,14] := -0.46343678;
      W_f[3,15] := 0.83569944;
      W_f[3,16] := -0.05430738;
      W_f[3,17] := 0.70786965;
      W_f[3,18] := 0.19876151;
      W_f[3,19] := -0.69915366;
      W_f[3,20] := -0.17611495;
      W_f[3,21] := 0.20092955;
      W_f[3,22] := -0.14438288;
      W_f[3,23] := -0.42021966;
      W_f[3,24] := -1.73890960;
      W_f[3,25] := -1.93748581;
      W_f[3,26] := 0.37437740;
      W_f[3,27] := -0.33648852;
      W_f[3,28] := -0.52998650;
      W_f[3,29] := -0.21540485;
      W_f[3,30] := 0.12346305;
      W_f[3,31] := -1.46652377;
      W_f[3,32] := -0.06444205;
      W_f[3,33] := -0.11098939;
      W_f[3,34] := -1.70861423;
      W_f[3,35] := 0.08646686;
      W_f[3,36] := -0.31241891;
      W_f[3,37] := 0.18405192;
      W_f[3,38] := 0.09597546;
      W_f[3,39] := -0.47231856;
      W_f[4,0] := -0.68655890;
      W_f[4,1] := -0.13217999;
      W_f[4,2] := 0.35625494;
      W_f[4,3] := 0.30554897;
      W_f[4,4] := -0.03162502;
      W_f[4,5] := -0.29792979;
      W_f[4,6] := 0.58917129;
      W_f[4,7] := -0.73093665;
      W_f[4,8] := 0.45340016;
      W_f[4,9] := -0.78049994;
      W_f[4,10] := 1.06470847;
      W_f[4,11] := -0.72154427;
      W_f[4,12] := 0.61361283;
      W_f[4,13] := -0.15808085;
      W_f[4,14] := 0.16161436;
      W_f[4,15] := 0.49596149;
      W_f[4,16] := 0.16095451;
      W_f[4,17] := -0.06179220;
      W_f[4,18] := 0.32785669;
      W_f[4,19] := -0.55550033;
      W_f[4,20] := 0.33831125;
      W_f[4,21] := 0.42008299;
      W_f[4,22] := 0.14018138;
      W_f[4,23] := 0.07146686;
      W_f[4,24] := -1.39041436;
      W_f[4,25] := -1.03200912;
      W_f[4,26] := -0.01316805;
      W_f[4,27] := -0.44839305;
      W_f[4,28] := 0.26812327;
      W_f[4,29] := 0.52243602;
      W_f[4,30] := 0.16244783;
      W_f[4,31] := 0.08064588;
      W_f[4,32] := 0.15116373;
      W_f[4,33] := 0.27706525;
      W_f[4,34] := 0.00838195;
      W_f[4,35] := 0.22120388;
      W_f[4,36] := 0.00388904;
      W_f[4,37] := 0.23256938;
      W_f[4,38] := 0.03672211;
      W_f[4,39] := -0.05871196;
      W_f[5,0] := -0.31850499;
      W_f[5,1] := -0.19392890;
      W_f[5,2] := 0.22627491;
      W_f[5,3] := 0.23169017;
      W_f[5,4] := -0.03339583;
      W_f[5,5] := -0.05071303;
      W_f[5,6] := -0.10622723;
      W_f[5,7] := -0.33521771;
      W_f[5,8] := -0.07157414;
      W_f[5,9] := -0.09234001;
      W_f[5,10] := -0.14189070;
      W_f[5,11] := -0.08683578;
      W_f[5,12] := -0.33746284;
      W_f[5,13] := 0.10314211;
      W_f[5,14] := 0.03929972;
      W_f[5,15] := -0.19532774;
      W_f[5,16] := -0.02381146;
      W_f[5,17] := -0.05064490;
      W_f[5,18] := 0.07619996;
      W_f[5,19] := 0.00605248;
      W_f[5,20] := -0.16619976;
      W_f[5,21] := -0.18192923;
      W_f[5,22] := -0.02836195;
      W_f[5,23] := -0.16396762;
      W_f[5,24] := 1.19843626;
      W_f[5,25] := 1.41340172;
      W_f[5,26] := -0.01094361;
      W_f[5,27] := 0.30434716;
      W_f[5,28] := 0.11668126;
      W_f[5,29] := -0.07706277;
      W_f[5,30] := -0.14868948;
      W_f[5,31] := -0.06208035;
      W_f[5,32] := -0.03129140;
      W_f[5,33] := 0.03850839;
      W_f[5,34] := 0.35154325;
      W_f[5,35] := -0.13979124;
      W_f[5,36] := 0.09827670;
      W_f[5,37] := -0.27274382;
      W_f[5,38] := 0.22190601;
      W_f[5,39] := -0.08572483;
      W_f[6,0] := 0.42435455;
      W_f[6,1] := 0.08249456;
      W_f[6,2] := -0.18963394;
      W_f[6,3] := 0.96772748;
      W_f[6,4] := -0.09344198;
      W_f[6,5] := 0.28461251;
      W_f[6,6] := 0.26882553;
      W_f[6,7] := 0.03824774;
      W_f[6,8] := -0.46005750;
      W_f[6,9] := -0.23360646;
      W_f[6,10] := -0.51570272;
      W_f[6,11] := 0.10533451;
      W_f[6,12] := -0.29385400;
      W_f[6,13] := 0.10406341;
      W_f[6,14] := -0.16624695;
      W_f[6,15] := -0.13436821;
      W_f[6,16] := 0.22478721;
      W_f[6,17] := -0.09131246;
      W_f[6,18] := 0.04823525;
      W_f[6,19] := 0.05260798;
      W_f[6,20] := -0.69891000;
      W_f[6,21] := 0.10713236;
      W_f[6,22] := 0.35655347;
      W_f[6,23] := 0.04896878;
      W_f[6,24] := 1.60622585;
      W_f[6,25] := 1.59777772;
      W_f[6,26] := 0.01397667;
      W_f[6,27] := 0.11062758;
      W_f[6,28] := -0.02002599;
      W_f[6,29] := -0.26235700;
      W_f[6,30] := 0.37919369;
      W_f[6,31] := 0.53207237;
      W_f[6,32] := 0.60770577;
      W_f[6,33] := 0.39742690;
      W_f[6,34] := 1.69826937;
      W_f[6,35] := 0.32700410;
      W_f[6,36] := 0.09589316;
      W_f[6,37] := 0.21720356;
      W_f[6,38] := 0.08525729;
      W_f[6,39] := -0.27763492;
      W_f[7,0] := 0.07349383;
      W_f[7,1] := 0.02822049;
      W_f[7,2] := -0.84481883;
      W_f[7,3] := -0.00570222;
      W_f[7,4] := -0.02442058;
      W_f[7,5] := 0.01488233;
      W_f[7,6] := -0.08660860;
      W_f[7,7] := 0.42620417;
      W_f[7,8] := -0.60038781;
      W_f[7,9] := 0.03975275;
      W_f[7,10] := -0.10148104;
      W_f[7,11] := 0.05718910;
      W_f[7,12] := -0.24106570;
      W_f[7,13] := -0.08941713;
      W_f[7,14] := 0.03560799;
      W_f[7,15] := -0.02408374;
      W_f[7,16] := -0.03861163;
      W_f[7,17] := 0.01301947;
      W_f[7,18] := 0.08077341;
      W_f[7,19] := -0.14269280;
      W_f[7,20] := -0.10094183;
      W_f[7,21] := -0.12904163;
      W_f[7,22] := 0.04183144;
      W_f[7,23] := 0.01284674;
      W_f[7,24] := -0.51689070;
      W_f[7,25] := -0.17367765;
      W_f[7,26] := -0.23541959;
      W_f[7,27] := 0.04862856;
      W_f[7,28] := 0.02250761;
      W_f[7,29] := 0.25177976;
      W_f[7,30] := -0.04562416;
      W_f[7,31] := 0.11538678;
      W_f[7,32] := 0.11963823;
      W_f[7,33] := -0.04533112;
      W_f[7,34] := -0.04678701;
      W_f[7,35] := 0.12872556;
      W_f[7,36] := -0.02270832;
      W_f[7,37] := -0.07886821;
      W_f[7,38] := 0.02381593;
      W_f[7,39] := 0.08858704;
      W_f[8,0] := -0.05206773;
      W_f[8,1] := 0.05427258;
      W_f[8,2] := 0.03702171;
      W_f[8,3] := -0.05017863;
      W_f[8,4] := 0.08655027;
      W_f[8,5] := 0.22196861;
      W_f[8,6] := 0.03162810;
      W_f[8,7] := 0.10221078;
      W_f[8,8] := 0.00455063;
      W_f[8,9] := 0.00628684;
      W_f[8,10] := -0.05337523;
      W_f[8,11] := 0.57790899;
      W_f[8,12] := -0.25566924;
      W_f[8,13] := 0.10859618;
      W_f[8,14] := -0.62317979;
      W_f[8,15] := -0.34060201;
      W_f[8,16] := 0.37791482;
      W_f[8,17] := 0.11984153;
      W_f[8,18] := 0.05718478;
      W_f[8,19] := -0.20448290;
      W_f[8,20] := -0.16286524;
      W_f[8,21] := 0.03390548;
      W_f[8,22] := 0.26846093;
      W_f[8,23] := 0.10364473;
      W_f[8,24] := 1.36088157;
      W_f[8,25] := 1.17845643;
      W_f[8,26] := -0.17945874;
      W_f[8,27] := -0.04318528;
      W_f[8,28] := 0.05277695;
      W_f[8,29] := 0.40008074;
      W_f[8,30] := 0.28982165;
      W_f[8,31] := 0.26548448;
      W_f[8,32] := 0.11699653;
      W_f[8,33] := -0.07936662;
      W_f[8,34] := 1.23291886;
      W_f[8,35] := -0.10220630;
      W_f[8,36] := 0.04077746;
      W_f[8,37] := -0.01109453;
      W_f[8,38] := -0.00270548;
      W_f[8,39] := 0.32922214;
      W_f[9,0] := 0.05573991;
      W_f[9,1] := 0.15928070;
      W_f[9,2] := -0.20538576;
      W_f[9,3] := -0.22553030;
      W_f[9,4] := 0.05168120;
      W_f[9,5] := 0.05359697;
      W_f[9,6] := 0.26185945;
      W_f[9,7] := -0.13908036;
      W_f[9,8] := 0.28974172;
      W_f[9,9] := 0.10875951;
      W_f[9,10] := 0.05757365;
      W_f[9,11] := -0.50996691;
      W_f[9,12] := 0.28445700;
      W_f[9,13] := -0.10266189;
      W_f[9,14] := 0.04574974;
      W_f[9,15] := 0.04567835;
      W_f[9,16] := -0.10557504;
      W_f[9,17] := -0.02136442;
      W_f[9,18] := 0.07768130;
      W_f[9,19] := 0.39294431;
      W_f[9,20] := 0.47319910;
      W_f[9,21] := 0.47894293;
      W_f[9,22] := 0.48117480;
      W_f[9,23] := -0.14602897;
      W_f[9,24] := -1.63407671;
      W_f[9,25] := -1.23110938;
      W_f[9,26] := 0.20508099;
      W_f[9,27] := -0.38148832;
      W_f[9,28] := -0.21609570;
      W_f[9,29] := 0.25101468;
      W_f[9,30] := 0.29295075;
      W_f[9,31] := 0.17286620;
      W_f[9,32] := -0.12084815;
      W_f[9,33] := -0.02219285;
      W_f[9,34] := 0.73441553;
      W_f[9,35] := 0.28961566;
      W_f[9,36] := 0.37668696;
      W_f[9,37] := 0.11451841;
      W_f[9,38] := 0.21723421;
      W_f[9,39] := -0.12171413;
      W_f[10,0] := 0.06705637;
      W_f[10,1] := 0.13236697;
      W_f[10,2] := -0.06536680;
      W_f[10,3] := -0.55446088;
      W_f[10,4] := -0.05074413;
      W_f[10,5] := 0.09033373;
      W_f[10,6] := -0.11670884;
      W_f[10,7] := 0.11099172;
      W_f[10,8] := -0.04687689;
      W_f[10,9] := 0.48866400;
      W_f[10,10] := 0.04315257;
      W_f[10,11] := -0.67770696;
      W_f[10,12] := 0.34806654;
      W_f[10,13] := -0.25238055;
      W_f[10,14] := -0.04166590;
      W_f[10,15] := -0.09219848;
      W_f[10,16] := 0.03033659;
      W_f[10,17] := 0.19120644;
      W_f[10,18] := -0.53988522;
      W_f[10,19] := 0.06212352;
      W_f[10,20] := 0.00374554;
      W_f[10,21] := 0.24568129;
      W_f[10,22] := -0.00730431;
      W_f[10,23] := 0.00483285;
      W_f[10,24] := -0.41010752;
      W_f[10,25] := -0.42264855;
      W_f[10,26] := -0.17979439;
      W_f[10,27] := -0.22658983;
      W_f[10,28] := 0.25472331;
      W_f[10,29] := 0.09937658;
      W_f[10,30] := -0.23006694;
      W_f[10,31] := -0.32560429;
      W_f[10,32] := -0.11242366;
      W_f[10,33] := 0.03228963;
      W_f[10,34] := -0.63356531;
      W_f[10,35] := 0.00331152;
      W_f[10,36] := -0.01774516;
      W_f[10,37] := 0.09553108;
      W_f[10,38] := -0.03525795;
      W_f[10,39] := 0.09118873;
      W_f[11,0] := -0.05548671;
      W_f[11,1] := 0.04312468;
      W_f[11,2] := 0.05087255;
      W_f[11,3] := -0.20145284;
      W_f[11,4] := -0.12363057;
      W_f[11,5] := 0.01457960;
      W_f[11,6] := 0.00399208;
      W_f[11,7] := -0.15979573;
      W_f[11,8] := 0.07721531;
      W_f[11,9] := 0.09382067;
      W_f[11,10] := 0.14348166;
      W_f[11,11] := 0.02369672;
      W_f[11,12] := 0.01268554;
      W_f[11,13] := 0.00390034;
      W_f[11,14] := -0.08125563;
      W_f[11,15] := -0.08493713;
      W_f[11,16] := -0.00230125;
      W_f[11,17] := 0.00543362;
      W_f[11,18] := 0.03282235;
      W_f[11,19] := 0.15100349;
      W_f[11,20] := 0.08062916;
      W_f[11,21] := 0.10192282;
      W_f[11,22] := -0.05395636;
      W_f[11,23] := 0.02045641;
      W_f[11,24] := -1.06981623;
      W_f[11,25] := -0.96444160;
      W_f[11,26] := 0.11357144;
      W_f[11,27] := -0.10241026;
      W_f[11,28] := 0.01148179;
      W_f[11,29] := 0.57609814;
      W_f[11,30] := 0.11210281;
      W_f[11,31] := 0.26540700;
      W_f[11,32] := 0.00766895;
      W_f[11,33] := 0.24361147;
      W_f[11,34] := -0.19100992;
      W_f[11,35] := 0.13836668;
      W_f[11,36] := -0.07907706;
      W_f[11,37] := 0.16210142;
      W_f[11,38] := -0.08032323;
      W_f[11,39] := 0.03944568;
      W_f[12,0] := -0.09712142;
      W_f[12,1] := 0.15042873;
      W_f[12,2] := 0.00185882;
      W_f[12,3] := 0.30617756;
      W_f[12,4] := -0.02837334;
      W_f[12,5] := 0.03159374;
      W_f[12,6] := 0.02653202;
      W_f[12,7] := -0.19543266;
      W_f[12,8] := -0.54019034;
      W_f[12,9] := 0.30703321;
      W_f[12,10] := 0.01940106;
      W_f[12,11] := -0.00073306;
      W_f[12,12] := -0.05447024;
      W_f[12,13] := 0.11511699;
      W_f[12,14] := 0.03176329;
      W_f[12,15] := -0.11075164;
      W_f[12,16] := 0.01435645;
      W_f[12,17] := 0.00481650;
      W_f[12,18] := -0.44951710;
      W_f[12,19] := -0.30256301;
      W_f[12,20] := 0.01976250;
      W_f[12,21] := 0.17333755;
      W_f[12,22] := 0.06146537;
      W_f[12,23] := -0.08121999;
      W_f[12,24] := -0.92103386;
      W_f[12,25] := -0.75615406;
      W_f[12,26] := -0.03370170;
      W_f[12,27] := 0.12443633;
      W_f[12,28] := 0.29289612;
      W_f[12,29] := 0.49214187;
      W_f[12,30] := 0.18102019;
      W_f[12,31] := 0.07411977;
      W_f[12,32] := -0.03247951;
      W_f[12,33] := 0.32056615;
      W_f[12,34] := -0.32351911;
      W_f[12,35] := 0.04861661;
      W_f[12,36] := -0.06008893;
      W_f[12,37] := 0.08359354;
      W_f[12,38] := 0.12238526;
      W_f[12,39] := -0.09088918;
      W_f[13,0] := -0.03996856;
      W_f[13,1] := -0.07003301;
      W_f[13,2] := 0.48738447;
      W_f[13,3] := 0.42322090;
      W_f[13,4] := 0.19929154;
      W_f[13,5] := -0.00825110;
      W_f[13,6] := -0.05568064;
      W_f[13,7] := -0.09145232;
      W_f[13,8] := -0.14745592;
      W_f[13,9] := -0.42382202;
      W_f[13,10] := -0.20620814;
      W_f[13,11] := 0.26426822;
      W_f[13,12] := 0.06960107;
      W_f[13,13] := 0.00838765;
      W_f[13,14] := -0.33020329;
      W_f[13,15] := -0.00234537;
      W_f[13,16] := 0.02060067;
      W_f[13,17] := -0.54517114;
      W_f[13,18] := -0.13411263;
      W_f[13,19] := -0.30789149;
      W_f[13,20] := -0.42978236;
      W_f[13,21] := -0.08678114;
      W_f[13,22] := 0.37233558;
      W_f[13,23] := -0.06351268;
      W_f[13,24] := 2.38407421;
      W_f[13,25] := 2.23805380;
      W_f[13,26] := -0.19631039;
      W_f[13,27] := 0.08246402;
      W_f[13,28] := -0.04395683;
      W_f[13,29] := -0.28599751;
      W_f[13,30] := 0.44259760;
      W_f[13,31] := 0.18553278;
      W_f[13,32] := 0.47523347;
      W_f[13,33] := 0.45066708;
      W_f[13,34] := 2.39121842;
      W_f[13,35] := 0.19777589;
      W_f[13,36] := 0.14772733;
      W_f[13,37] := 0.17772952;
      W_f[13,38] := -0.06637986;
      W_f[13,39] := 0.27313134;
      W_f[14,0] := -0.10999595;
      W_f[14,1] := 0.16378450;
      W_f[14,2] := 0.31294572;
      W_f[14,3] := 0.30457804;
      W_f[14,4] := 0.39332005;
      W_f[14,5] := 0.29185969;
      W_f[14,6] := 0.49079815;
      W_f[14,7] := 0.10466534;
      W_f[14,8] := -0.10972983;
      W_f[14,9] := -0.30818820;
      W_f[14,10] := -0.92225468;
      W_f[14,11] := -0.63368195;
      W_f[14,12] := 0.26334706;
      W_f[14,13] := -0.33846161;
      W_f[14,14] := 0.10465050;
      W_f[14,15] := -0.03916458;
      W_f[14,16] := 0.14926721;
      W_f[14,17] := 0.03337602;
      W_f[14,18] := -0.00833549;
      W_f[14,19] := 0.29542312;
      W_f[14,20] := 0.07174528;
      W_f[14,21] := 0.51826459;
      W_f[14,22] := 0.18384574;
      W_f[14,23] := 0.03958815;
      W_f[14,24] := -1.07650769;
      W_f[14,25] := -0.76949328;
      W_f[14,26] := 0.46225747;
      W_f[14,27] := -0.32431909;
      W_f[14,28] := -0.20283256;
      W_f[14,29] := 0.67629284;
      W_f[14,30] := 0.17858230;
      W_f[14,31] := 0.26788053;
      W_f[14,32] := 0.01443615;
      W_f[14,33] := 0.09308545;
      W_f[14,34] := 0.21026219;
      W_f[14,35] := -0.08981100;
      W_f[14,36] := -0.13266245;
      W_f[14,37] := -0.12135204;
      W_f[14,38] := -0.21469142;
      W_f[14,39] := -0.25131592;
      W_f[15,0] := -0.16556653;
      W_f[15,1] := -0.06627338;
      W_f[15,2] := 0.04116353;
      W_f[15,3] := -0.30215326;
      W_f[15,4] := 0.12548773;
      W_f[15,5] := 0.16821291;
      W_f[15,6] := -0.22060153;
      W_f[15,7] := -0.06172123;
      W_f[15,8] := 0.04885555;
      W_f[15,9] := 0.02473416;
      W_f[15,10] := -0.03054220;
      W_f[15,11] := 0.15292585;
      W_f[15,12] := 0.00023254;
      W_f[15,13] := -0.00098793;
      W_f[15,14] := -0.07777366;
      W_f[15,15] := -0.18486318;
      W_f[15,16] := -0.02031197;
      W_f[15,17] := 0.08086631;
      W_f[15,18] := -0.01069839;
      W_f[15,19] := 0.05074516;
      W_f[15,20] := 0.15063727;
      W_f[15,21] := 0.01365798;
      W_f[15,22] := 0.13210511;
      W_f[15,23] := -0.05615190;
      W_f[15,24] := -0.92742151;
      W_f[15,25] := -0.65037620;
      W_f[15,26] := 0.01558890;
      W_f[15,27] := 0.18203004;
      W_f[15,28] := 0.03965090;
      W_f[15,29] := -0.07643162;
      W_f[15,30] := 0.02053319;
      W_f[15,31] := 0.12344345;
      W_f[15,32] := 0.35255781;
      W_f[15,33] := 0.31968316;
      W_f[15,34] := 0.22691649;
      W_f[15,35] := 0.09319179;
      W_f[15,36] := 0.09234352;
      W_f[15,37] := -0.16712017;
      W_f[15,38] := -0.04719787;
      W_f[15,39] := 0.65844274;
      W_f[16,0] := 0.22374457;
      W_f[16,1] := 0.05910943;
      W_f[16,2] := -0.06322084;
      W_f[16,3] := 0.27774197;
      W_f[16,4] := -0.13294286;
      W_f[16,5] := -0.14119923;
      W_f[16,6] := -0.26860869;
      W_f[16,7] := 0.15995319;
      W_f[16,8] := 0.02333695;
      W_f[16,9] := -0.17028902;
      W_f[16,10] := 0.22073960;
      W_f[16,11] := -0.76096177;
      W_f[16,12] := -0.48183411;
      W_f[16,13] := 0.32877094;
      W_f[16,14] := 0.38851735;
      W_f[16,15] := -0.30537850;
      W_f[16,16] := -0.12814270;
      W_f[16,17] := -0.39573076;
      W_f[16,18] := 0.18768115;
      W_f[16,19] := 0.52345359;
      W_f[16,20] := -0.35657167;
      W_f[16,21] := -0.27201805;
      W_f[16,22] := -0.11477985;
      W_f[16,23] := -0.31365654;
      W_f[16,24] := 0.08666131;
      W_f[16,25] := 0.21089429;
      W_f[16,26] := -0.11963987;
      W_f[16,27] := -0.12481143;
      W_f[16,28] := 0.10807389;
      W_f[16,29] := -0.17113568;
      W_f[16,30] := -0.35757676;
      W_f[16,31] := 0.36995792;
      W_f[16,32] := -0.18190899;
      W_f[16,33] := 0.16161774;
      W_f[16,34] := -0.24879223;
      W_f[16,35] := -0.08751137;
      W_f[16,36] := -0.04311307;
      W_f[16,37] := -0.17220454;
      W_f[16,38] := 0.19482853;
      W_f[16,39] := -0.16588378;
      W_f[17,0] := -0.16411990;
      W_f[17,1] := 0.09834433;
      W_f[17,2] := 0.25410935;
      W_f[17,3] := 0.40745008;
      W_f[17,4] := -0.15107033;
      W_f[17,5] := 0.23475306;
      W_f[17,6] := -0.24045940;
      W_f[17,7] := 0.10921574;
      W_f[17,8] := -0.17072932;
      W_f[17,9] := -0.08083232;
      W_f[17,10] := -0.18766029;
      W_f[17,11] := -0.33869505;
      W_f[17,12] := 0.17434444;
      W_f[17,13] := 0.01097766;
      W_f[17,14] := 0.16010438;
      W_f[17,15] := -0.05596434;
      W_f[17,16] := 0.10686168;
      W_f[17,17] := 0.12036951;
      W_f[17,18] := 0.16494197;
      W_f[17,19] := 0.12652035;
      W_f[17,20] := -0.00716413;
      W_f[17,21] := 0.36908007;
      W_f[17,22] := 0.21722621;
      W_f[17,23] := -0.00221541;
      W_f[17,24] := -0.33342555;
      W_f[17,25] := -0.46759641;
      W_f[17,26] := -0.06185902;
      W_f[17,27] := -0.21750233;
      W_f[17,28] := 0.22360668;
      W_f[17,29] := 0.09053066;
      W_f[17,30] := 0.09899973;
      W_f[17,31] := -0.08313378;
      W_f[17,32] := 0.32378528;
      W_f[17,33] := 0.20052801;
      W_f[17,34] := -1.02485752;
      W_f[17,35] := 0.03071750;
      W_f[17,36] := 0.01856773;
      W_f[17,37] := 0.12227248;
      W_f[17,38] := 0.02499303;
      W_f[17,39] := -0.81374878;
      W_f[18,0] := 0.36294127;
      W_f[18,1] := 0.02575219;
      W_f[18,2] := -0.17604761;
      W_f[18,3] := -0.33789763;
      W_f[18,4] := -0.07201187;
      W_f[18,5] := 0.08762357;
      W_f[18,6] := -0.23841025;
      W_f[18,7] := 0.19438463;
      W_f[18,8] := -0.10556871;
      W_f[18,9] := -0.15092371;
      W_f[18,10] := 0.10175239;
      W_f[18,11] := 0.11924792;
      W_f[18,12] := -0.14140444;
      W_f[18,13] := 0.02214300;
      W_f[18,14] := 0.17515695;
      W_f[18,15] := -0.06727323;
      W_f[18,16] := 0.22449253;
      W_f[18,17] := -0.01732972;
      W_f[18,18] := -0.00555121;
      W_f[18,19] := -0.19859479;
      W_f[18,20] := -0.14399439;
      W_f[18,21] := 0.09881490;
      W_f[18,22] := 0.10322018;
      W_f[18,23] := -0.03669460;
      W_f[18,24] := -0.73212147;
      W_f[18,25] := -0.60783029;
      W_f[18,26] := 0.07082136;
      W_f[18,27] := -0.09695113;
      W_f[18,28] := 0.02489661;
      W_f[18,29] := -0.26595870;
      W_f[18,30] := 0.12078937;
      W_f[18,31] := -0.88141137;
      W_f[18,32] := 0.01366802;
      W_f[18,33] := -0.30026230;
      W_f[18,34] := -0.01247005;
      W_f[18,35] := 0.16910952;
      W_f[18,36] := -0.25617203;
      W_f[18,37] := 0.15913877;
      W_f[18,38] := -0.07596558;
      W_f[18,39] := -0.16493645;
      W_f[19,0] := -0.01734783;
      W_f[19,1] := 0.13046260;
      W_f[19,2] := -0.14956820;
      W_f[19,3] := -0.13372861;
      W_f[19,4] := 0.01607699;
      W_f[19,5] := -0.03008930;
      W_f[19,6] := -0.03232536;
      W_f[19,7] := 0.13831176;
      W_f[19,8] := 0.05940061;
      W_f[19,9] := -0.13088953;
      W_f[19,10] := 0.01243817;
      W_f[19,11] := -0.17900078;
      W_f[19,12] := 0.29835901;
      W_f[19,13] := 0.30771545;
      W_f[19,14] := -0.08315364;
      W_f[19,15] := -0.32168353;
      W_f[19,16] := 0.32334423;
      W_f[19,17] := -0.04730310;
      W_f[19,18] := 0.09356403;
      W_f[19,19] := 0.52750629;
      W_f[19,20] := 0.06653363;
      W_f[19,21] := 0.20962518;
      W_f[19,22] := 0.29950517;
      W_f[19,23] := -0.19698098;
      W_f[19,24] := 0.20843033;
      W_f[19,25] := 0.66837531;
      W_f[19,26] := -0.11612438;
      W_f[19,27] := -0.26898244;
      W_f[19,28] := 0.03650144;
      W_f[19,29] := -0.16495816;
      W_f[19,30] := 0.25047439;
      W_f[19,31] := -0.00991298;
      W_f[19,32] := -0.05104885;
      W_f[19,33] := 0.10937680;
      W_f[19,34] := -0.67745608;
      W_f[19,35] := 0.10768792;
      W_f[19,36] := 0.11150705;
      W_f[19,37] := 0.00372975;
      W_f[19,38] := -0.40008494;
      W_f[19,39] := 0.45059848;
      W_f[20,0] := 0.05295354;
      W_f[20,1] := -0.13710082;
      W_f[20,2] := -0.12655978;
      W_f[20,3] := -0.52311695;
      W_f[20,4] := 0.10019384;
      W_f[20,5] := 0.12332516;
      W_f[20,6] := -0.04756395;
      W_f[20,7] := 0.06900418;
      W_f[20,8] := -0.83848727;
      W_f[20,9] := 1.02468872;
      W_f[20,10] := -0.20606503;
      W_f[20,11] := 0.19898677;
      W_f[20,12] := -0.13268803;
      W_f[20,13] := 0.03680019;
      W_f[20,14] := 0.01324347;
      W_f[20,15] := 0.05220984;
      W_f[20,16] := 0.22231728;
      W_f[20,17] := 0.05803931;
      W_f[20,18] := -0.15821685;
      W_f[20,19] := -0.18480341;
      W_f[20,20] := -0.11115044;
      W_f[20,21] := -0.04297195;
      W_f[20,22] := 0.31193075;
      W_f[20,23] := -0.03074704;
      W_f[20,24] := 1.41226840;
      W_f[20,25] := 1.53308392;
      W_f[20,26] := 0.05630440;
      W_f[20,27] := 0.05454231;
      W_f[20,28] := -0.23422292;
      W_f[20,29] := -0.21086636;
      W_f[20,30] := 0.45930535;
      W_f[20,31] := 0.09115323;
      W_f[20,32] := 0.05492384;
      W_f[20,33] := 0.00805198;
      W_f[20,34] := 1.54443157;
      W_f[20,35] := -0.01436506;
      W_f[20,36] := -0.17954412;
      W_f[20,37] := -0.09542100;
      W_f[20,38] := 0.24947862;
      W_f[20,39] := -0.10104286;
      W_f[21,0] := -0.00168017;
      W_f[21,1] := 0.11660825;
      W_f[21,2] := -0.00404962;
      W_f[21,3] := 0.36214161;
      W_f[21,4] := 0.34586513;
      W_f[21,5] := 0.06963939;
      W_f[21,6] := -0.00849801;
      W_f[21,7] := -0.10223118;
      W_f[21,8] := -0.10811724;
      W_f[21,9] := 0.04582016;
      W_f[21,10] := -0.26858315;
      W_f[21,11] := 0.40021136;
      W_f[21,12] := 0.00788286;
      W_f[21,13] := -0.07432951;
      W_f[21,14] := 0.05539732;
      W_f[21,15] := 0.02197883;
      W_f[21,16] := 0.28201821;
      W_f[21,17] := -0.21401763;
      W_f[21,18] := -0.29455173;
      W_f[21,19] := -0.04343071;
      W_f[21,20] := -0.11677518;
      W_f[21,21] := -0.40573204;
      W_f[21,22] := 0.34463850;
      W_f[21,23] := 0.02065710;
      W_f[21,24] := 0.62987918;
      W_f[21,25] := 0.62826115;
      W_f[21,26] := -0.16319363;
      W_f[21,27] := 0.35674879;
      W_f[21,28] := -0.02922228;
      W_f[21,29] := 0.63345420;
      W_f[21,30] := 0.23994400;
      W_f[21,31] := 0.06582332;
      W_f[21,32] := 0.20053940;
      W_f[21,33] := 0.05011126;
      W_f[21,34] := 0.13510664;
      W_f[21,35] := 0.36979461;
      W_f[21,36] := 0.30219561;
      W_f[21,37] := 0.36491936;
      W_f[21,38] := 0.08422065;
      W_f[21,39] := 0.28683770;
      W_f[22,0] := -0.59764260;
      W_f[22,1] := 0.11420204;
      W_f[22,2] := 0.49944505;
      W_f[22,3] := -0.16634117;
      W_f[22,4] := 0.13442634;
      W_f[22,5] := -0.05985187;
      W_f[22,6] := 0.17724130;
      W_f[22,7] := 0.13804770;
      W_f[22,8] := -0.24538754;
      W_f[22,9] := 0.21552241;
      W_f[22,10] := 0.14287704;
      W_f[22,11] := -0.12601700;
      W_f[22,12] := 0.26320851;
      W_f[22,13] := 0.16650802;
      W_f[22,14] := -0.21341632;
      W_f[22,15] := -0.54411554;
      W_f[22,16] := 0.30557558;
      W_f[22,17] := -0.22573556;
      W_f[22,18] := -1.05107760;
      W_f[22,19] := 0.29967535;
      W_f[22,20] := -0.08190977;
      W_f[22,21] := 0.09606460;
      W_f[22,22] := -0.34405023;
      W_f[22,23] := -0.40458128;
      W_f[22,24] := -0.40848887;
      W_f[22,25] := -0.39460698;
      W_f[22,26] := 0.21953718;
      W_f[22,27] := -0.08266225;
      W_f[22,28] := -0.21698205;
      W_f[22,29] := 0.33896431;
      W_f[22,30] := -0.31644160;
      W_f[22,31] := -0.82518321;
      W_f[22,32] := -0.13789199;
      W_f[22,33] := -0.06215421;
      W_f[22,34] := -0.24466747;
      W_f[22,35] := 0.18926638;
      W_f[22,36] := -0.07384060;
      W_f[22,37] := 0.36008319;
      W_f[22,38] := -0.16622342;
      W_f[22,39] := -0.12244521;
      W_f[23,0] := 0.10097027;
      W_f[23,1] := -0.13139288;
      W_f[23,2] := -0.14940387;
      W_f[23,3] := -0.24939288;
      W_f[23,4] := 0.09224908;
      W_f[23,5] := 0.02639719;
      W_f[23,6] := -0.20195131;
      W_f[23,7] := -0.01629142;
      W_f[23,8] := 0.41546646;
      W_f[23,9] := 0.50435215;
      W_f[23,10] := -0.38946828;
      W_f[23,11] := 0.14280544;
      W_f[23,12] := -0.26078326;
      W_f[23,13] := 0.13182658;
      W_f[23,14] := -0.15221739;
      W_f[23,15] := -0.32292679;
      W_f[23,16] := 0.09519158;
      W_f[23,17] := -0.10446651;
      W_f[23,18] := 0.11899559;
      W_f[23,19] := -0.44001421;
      W_f[23,20] := 0.02194781;
      W_f[23,21] := -0.26942325;
      W_f[23,22] := 0.03859116;
      W_f[23,23] := 0.04861640;
      W_f[23,24] := -0.29334232;
      W_f[23,25] := -0.39534897;
      W_f[23,26] := -0.19794963;
      W_f[23,27] := 0.54521793;
      W_f[23,28] := 0.07424716;
      W_f[23,29] := -0.18977107;
      W_f[23,30] := 0.06721469;
      W_f[23,31] := -0.09336343;
      W_f[23,32] := -0.03395103;
      W_f[23,33] := -0.16725579;
      W_f[23,34] := 0.01551263;
      W_f[23,35] := -0.13205801;
      W_f[23,36] := -0.04547273;
      W_f[23,37] := 0.17488526;
      W_f[23,38] := 0.08316690;
      W_f[23,39] := -0.08328584;
      W_f[24,0] := 0.13098057;
      W_f[24,1] := -0.06250014;
      W_f[24,2] := -0.00119376;
      W_f[24,3] := -0.07479530;
      W_f[24,4] := -0.18538533;
      W_f[24,5] := -0.01275790;
      W_f[24,6] := 0.00874758;
      W_f[24,7] := 0.12383805;
      W_f[24,8] := -0.04926819;
      W_f[24,9] := -0.01701698;
      W_f[24,10] := -0.06444911;
      W_f[24,11] := 0.21160479;
      W_f[24,12] := -0.02235752;
      W_f[24,13] := 0.00378762;
      W_f[24,14] := 0.02738534;
      W_f[24,15] := 0.17725867;
      W_f[24,16] := -0.19304124;
      W_f[24,17] := -0.01714083;
      W_f[24,18] := -0.01785743;
      W_f[24,19] := -0.62033468;
      W_f[24,20] := -0.12589391;
      W_f[24,21] := -0.39348763;
      W_f[24,22] := 0.31992048;
      W_f[24,23] := -0.27218062;
      W_f[24,24] := 1.81270516;
      W_f[24,25] := 1.65550554;
      W_f[24,26] := -0.26350173;
      W_f[24,27] := 0.06742683;
      W_f[24,28] := -0.11887355;
      W_f[24,29] := 0.43823522;
      W_f[24,30] := 0.17323317;
      W_f[24,31] := 0.32686615;
      W_f[24,32] := 0.37364411;
      W_f[24,33] := 0.15626027;
      W_f[24,34] := 1.55385089;
      W_f[24,35] := 0.28087455;
      W_f[24,36] := -0.18218301;
      W_f[24,37] := 0.42226493;
      W_f[24,38] := 0.08549567;
      W_f[24,39] := 0.47081169;
      W_f[25,0] := -0.05556887;
      W_f[25,1] := -0.03406537;
      W_f[25,2] := 0.14011057;
      W_f[25,3] := 0.14114504;
      W_f[25,4] := 0.00227548;
      W_f[25,5] := 0.12053847;
      W_f[25,6] := -0.05779338;
      W_f[25,7] := -0.22579378;
      W_f[25,8] := -0.06333803;
      W_f[25,9] := -0.00101634;
      W_f[25,10] := -0.11495918;
      W_f[25,11] := -0.05879531;
      W_f[25,12] := 0.04155201;
      W_f[25,13] := 0.03228154;
      W_f[25,14] := -0.37705407;
      W_f[25,15] := -0.53819382;
      W_f[25,16] := -0.13453944;
      W_f[25,17] := 0.27555528;
      W_f[25,18] := 0.01666597;
      W_f[25,19] := -0.22168976;
      W_f[25,20] := 0.05109134;
      W_f[25,21] := -0.00183230;
      W_f[25,22] := -0.01646283;
      W_f[25,23] := -0.02016181;
      W_f[25,24] := 0.73902524;
      W_f[25,25] := 0.93939823;
      W_f[25,26] := -0.08844233;
      W_f[25,27] := 0.04351176;
      W_f[25,28] := -0.03928512;
      W_f[25,29] := -0.01265163;
      W_f[25,30] := 0.14475761;
      W_f[25,31] := -0.10781216;
      W_f[25,32] := 0.18317719;
      W_f[25,33] := 0.33000368;
      W_f[25,34] := -0.57851905;
      W_f[25,35] := -0.09157128;
      W_f[25,36] := 0.09818074;
      W_f[25,37] := -0.18664096;
      W_f[25,38] := 0.04246709;
      W_f[25,39] := 0.07847621;
      W_f[26,0] := 0.14105089;
      W_f[26,1] := 0.09353172;
      W_f[26,2] := -0.33030543;
      W_f[26,3] := 0.43264621;
      W_f[26,4] := 0.24365731;
      W_f[26,5] := -0.11344527;
      W_f[26,6] := 0.03489910;
      W_f[26,7] := -0.34441987;
      W_f[26,8] := -0.24129467;
      W_f[26,9] := -0.26754951;
      W_f[26,10] := -0.13237664;
      W_f[26,11] := -0.25729531;
      W_f[26,12] := -0.18069156;
      W_f[26,13] := -0.01574439;
      W_f[26,14] := -0.29478207;
      W_f[26,15] := -0.82912469;
      W_f[26,16] := -0.12289927;
      W_f[26,17] := -0.31922388;
      W_f[26,18] := 0.09471790;
      W_f[26,19] := -0.13924044;
      W_f[26,20] := -0.23671141;
      W_f[26,21] := 0.14164712;
      W_f[26,22] := -0.03585915;
      W_f[26,23] := 0.96720719;
      W_f[26,24] := 0.72606045;
      W_f[26,25] := 0.50532269;
      W_f[26,26] := -0.29200366;
      W_f[26,27] := 0.19223879;
      W_f[26,28] := 0.09991259;
      W_f[26,29] := -0.09034248;
      W_f[26,30] := -0.00482521;
      W_f[26,31] := -0.11174250;
      W_f[26,32] := -0.09373572;
      W_f[26,33] := -0.00918921;
      W_f[26,34] := -0.26856694;
      W_f[26,35] := -0.16221951;
      W_f[26,36] := -0.02910131;
      W_f[26,37] := -0.09744545;
      W_f[26,38] := -0.03827441;
      W_f[26,39] := 0.35593715;
      W_f[27,0] := 0.06162736;
      W_f[27,1] := -0.00079178;
      W_f[27,2] := -0.45381555;
      W_f[27,3] := 0.06428052;
      W_f[27,4] := 0.04040126;
      W_f[27,5] := 0.12687680;
      W_f[27,6] := -0.00780606;
      W_f[27,7] := -0.10548334;
      W_f[27,8] := -0.19921654;
      W_f[27,9] := 0.23297761;
      W_f[27,10] := 0.06463186;
      W_f[27,11] := 0.03318268;
      W_f[27,12] := -0.03947852;
      W_f[27,13] := -0.00685048;
      W_f[27,14] := -0.00737523;
      W_f[27,15] := -0.21209772;
      W_f[27,16] := 0.45497540;
      W_f[27,17] := -0.36895815;
      W_f[27,18] := 0.15872858;
      W_f[27,19] := 0.44276521;
      W_f[27,20] := 0.00021969;
      W_f[27,21] := 0.17368497;
      W_f[27,22] := 0.20000930;
      W_f[27,23] := -0.08216770;
      W_f[27,24] := 0.78227371;
      W_f[27,25] := 0.88182676;
      W_f[27,26] := 0.00509356;
      W_f[27,27] := -0.07620359;
      W_f[27,28] := 0.05403636;
      W_f[27,29] := -0.18912379;
      W_f[27,30] := 0.34674552;
      W_f[27,31] := 0.04280552;
      W_f[27,32] := 0.21729645;
      W_f[27,33] := -0.09554624;
      W_f[27,34] := 0.61564386;
      W_f[27,35] := -0.03573473;
      W_f[27,36] := -0.05912105;
      W_f[27,37] := 0.20100754;
      W_f[27,38] := 0.14946508;
      W_f[27,39] := -0.08973806;
      W_f[28,0] := 0.08568294;
      W_f[28,1] := 0.07220396;
      W_f[28,2] := -0.00819603;
      W_f[28,3] := -0.48418882;
      W_f[28,4] := -0.11894052;
      W_f[28,5] := -0.02794145;
      W_f[28,6] := 0.12426823;
      W_f[28,7] := 0.30004731;
      W_f[28,8] := 0.05287009;
      W_f[28,9] := 0.00921909;
      W_f[28,10] := 0.00668684;
      W_f[28,11] := 0.06600591;
      W_f[28,12] := 0.25218466;
      W_f[28,13] := -0.16467427;
      W_f[28,14] := 0.00648815;
      W_f[28,15] := -0.00700287;
      W_f[28,16] := -0.11720763;
      W_f[28,17] := -0.02515974;
      W_f[28,18] := -0.00833579;
      W_f[28,19] := -0.03406101;
      W_f[28,20] := 0.07821744;
      W_f[28,21] := 0.03123923;
      W_f[28,22] := 0.12632163;
      W_f[28,23] := -0.04973659;
      W_f[28,24] := 0.09309764;
      W_f[28,25] := 0.26760951;
      W_f[28,26] := 0.05048810;
      W_f[28,27] := -0.16696256;
      W_f[28,28] := 0.03711645;
      W_f[28,29] := 0.33228141;
      W_f[28,30] := 0.12719348;
      W_f[28,31] := -0.02180708;
      W_f[28,32] := -0.04254036;
      W_f[28,33] := 0.29769444;
      W_f[28,34] := 0.00704242;
      W_f[28,35] := 0.17184366;
      W_f[28,36] := -0.01311863;
      W_f[28,37] := 0.04687236;
      W_f[28,38] := 0.09186333;
      W_f[28,39] := 0.06206822;
      W_f[29,0] := -0.29772484;
      W_f[29,1] := -0.06461336;
      W_f[29,2] := 0.26568708;
      W_f[29,3] := 0.08998085;
      W_f[29,4] := -0.05701882;
      W_f[29,5] := 0.22950536;
      W_f[29,6] := -0.05952236;
      W_f[29,7] := -0.47861040;
      W_f[29,8] := 0.43492243;
      W_f[29,9] := -0.07213128;
      W_f[29,10] := -0.03874899;
      W_f[29,11] := -0.03404453;
      W_f[29,12] := -0.15405726;
      W_f[29,13] := -0.48577595;
      W_f[29,14] := -0.02204370;
      W_f[29,15] := -0.05456595;
      W_f[29,16] := 0.05162636;
      W_f[29,17] := 0.02018623;
      W_f[29,18] := 0.49756289;
      W_f[29,19] := 0.03590911;
      W_f[29,20] := -0.17447828;
      W_f[29,21] := -0.24529612;
      W_f[29,22] := 0.06076729;
      W_f[29,23] := 0.02893092;
      W_f[29,24] := -0.28510767;
      W_f[29,25] := -0.37744424;
      W_f[29,26] := 0.11913476;
      W_f[29,27] := 0.08534627;
      W_f[29,28] := 0.14223781;
      W_f[29,29] := 0.04189867;
      W_f[29,30] := -0.11465988;
      W_f[29,31] := -0.11025470;
      W_f[29,32] := -0.05296186;
      W_f[29,33] := 0.05677674;
      W_f[29,34] := -0.11102781;
      W_f[29,35] := -0.10578488;
      W_f[29,36] := -0.42032716;
      W_f[29,37] := 0.17246746;
      W_f[29,38] := 0.08812485;
      W_f[29,39] := 0.46797311;
      W_f[30,0] := 0.02389588;
      W_f[30,1] := 0.03138966;
      W_f[30,2] := -0.07268680;
      W_f[30,3] := -0.47570822;
      W_f[30,4] := -0.01275609;
      W_f[30,5] := 0.06347569;
      W_f[30,6] := -0.11336186;
      W_f[30,7] := 0.19684200;
      W_f[30,8] := -0.16061504;
      W_f[30,9] := 0.33959588;
      W_f[30,10] := -0.08797532;
      W_f[30,11] := -0.02474829;
      W_f[30,12] := -0.01200104;
      W_f[30,13] := -0.04101486;
      W_f[30,14] := -0.00347323;
      W_f[30,15] := 0.27267310;
      W_f[30,16] := 0.12974751;
      W_f[30,17] := -0.13578549;
      W_f[30,18] := -0.00819293;
      W_f[30,19] := 0.19127662;
      W_f[30,20] := -0.01524954;
      W_f[30,21] := 0.05541044;
      W_f[30,22] := 0.17716034;
      W_f[30,23] := 0.02053385;
      W_f[30,24] := 0.26789400;
      W_f[30,25] := 0.29255810;
      W_f[30,26] := -0.12997754;
      W_f[30,27] := 0.04716227;
      W_f[30,28] := 0.12676223;
      W_f[30,29] := -0.20882915;
      W_f[30,30] := 0.22658019;
      W_f[30,31] := 0.21638000;
      W_f[30,32] := 0.06398591;
      W_f[30,33] := -0.08813185;
      W_f[30,34] := 0.69014442;
      W_f[30,35] := -0.20874223;
      W_f[30,36] := -0.03230392;
      W_f[30,37] := -0.09084769;
      W_f[30,38] := 0.21777090;
      W_f[30,39] := -0.12998870;
      W_f[31,0] := 0.25092110;
      W_f[31,1] := 0.91395742;
      W_f[31,2] := 0.01737494;
      W_f[31,3] := 0.17552799;
      W_f[31,4] := 0.00730009;
      W_f[31,5] := 0.29924333;
      W_f[31,6] := -0.13413790;
      W_f[31,7] := 0.44026881;
      W_f[31,8] := -0.06399131;
      W_f[31,9] := 0.16534172;
      W_f[31,10] := -0.21947183;
      W_f[31,11] := -0.08995450;
      W_f[31,12] := -0.00483328;
      W_f[31,13] := -0.09211861;
      W_f[31,14] := 0.20189485;
      W_f[31,15] := 0.03910992;
      W_f[31,16] := -0.38301164;
      W_f[31,17] := 0.16348492;
      W_f[31,18] := -0.02939895;
      W_f[31,19] := -0.42179126;
      W_f[31,20] := 0.18242118;
      W_f[31,21] := 0.45759532;
      W_f[31,22] := 0.00682034;
      W_f[31,23] := -0.09145424;
      W_f[31,24] := 1.18018579;
      W_f[31,25] := 1.11625838;
      W_f[31,26] := -0.26431102;
      W_f[31,27] := -0.07003646;
      W_f[31,28] := 0.15999524;
      W_f[31,29] := 0.26074442;
      W_f[31,30] := 0.17888932;
      W_f[31,31] := 0.08699726;
      W_f[31,32] := 0.18072855;
      W_f[31,33] := 0.13479882;
      W_f[31,34] := 0.10072931;
      W_f[31,35] := -0.20896043;
      W_f[31,36] := 0.00694057;
      W_f[31,37] := -0.12319652;
      W_f[31,38] := 0.39178091;
      W_f[31,39] := -0.17493194;
      W_g[0,0] := -0.05221632;
      W_g[0,1] := 0.07101889;
      W_g[0,2] := -0.22668254;
      W_g[0,3] := -0.06343202;
      W_g[0,4] := -0.34505597;
      W_g[0,5] := 0.02013769;
      W_g[0,6] := 0.13723709;
      W_g[0,7] := 0.01286843;
      W_g[0,8] := 0.25928411;
      W_g[0,9] := 0.15451054;
      W_g[0,10] := -0.01147146;
      W_g[0,11] := -0.14489363;
      W_g[0,12] := -0.09124152;
      W_g[0,13] := -0.16375518;
      W_g[0,14] := 0.00021868;
      W_g[0,15] := -0.18328460;
      W_g[0,16] := 0.00898300;
      W_g[0,17] := -0.14367449;
      W_g[0,18] := -0.02342481;
      W_g[0,19] := -0.03811495;
      W_g[0,20] := 0.38238192;
      W_g[0,21] := -0.33150980;
      W_g[0,22] := -0.11630447;
      W_g[0,23] := 0.17661096;
      W_g[0,24] := 0.37532377;
      W_g[0,25] := 0.47437796;
      W_g[0,26] := 0.30349693;
      W_g[0,27] := 0.39895791;
      W_g[0,28] := 0.33480498;
      W_g[0,29] := -0.04643648;
      W_g[0,30] := -0.13288611;
      W_g[0,31] := 0.12894422;
      W_g[0,32] := 0.02159341;
      W_g[0,33] := 0.02643129;
      W_g[0,34] := 0.54021758;
      W_g[0,35] := 0.08358868;
      W_g[0,36] := 0.05316209;
      W_g[0,37] := 0.13387355;
      W_g[0,38] := 0.05129709;
      W_g[0,39] := -0.18220155;
      W_g[1,0] := 0.11506090;
      W_g[1,1] := 0.13651496;
      W_g[1,2] := 0.05378669;
      W_g[1,3] := 0.23183541;
      W_g[1,4] := 0.31218642;
      W_g[1,5] := 1.26320171;
      W_g[1,6] := 0.57657862;
      W_g[1,7] := 0.48835528;
      W_g[1,8] := -0.11248570;
      W_g[1,9] := 0.39191779;
      W_g[1,10] := 0.36195213;
      W_g[1,11] := -0.06714219;
      W_g[1,12] := -0.22399405;
      W_g[1,13] := 0.29271981;
      W_g[1,14] := -0.01325159;
      W_g[1,15] := 0.02355744;
      W_g[1,16] := 0.02834371;
      W_g[1,17] := -0.00796816;
      W_g[1,18] := 0.05731512;
      W_g[1,19] := 0.00908184;
      W_g[1,20] := 0.46170649;
      W_g[1,21] := 0.16210626;
      W_g[1,22] := 0.00231385;
      W_g[1,23] := -0.02824998;
      W_g[1,24] := 0.04692646;
      W_g[1,25] := 0.07125357;
      W_g[1,26] := -0.05206983;
      W_g[1,27] := -0.06304284;
      W_g[1,28] := -0.05542786;
      W_g[1,29] := 0.12507403;
      W_g[1,30] := 0.15066417;
      W_g[1,31] := -0.00473702;
      W_g[1,32] := 0.00781616;
      W_g[1,33] := -0.04659111;
      W_g[1,34] := -0.01626356;
      W_g[1,35] := -0.04343637;
      W_g[1,36] := -0.05985352;
      W_g[1,37] := 0.06222189;
      W_g[1,38] := 0.03715008;
      W_g[1,39] := 0.06825569;
      W_g[2,0] := 0.17983484;
      W_g[2,1] := -0.37871104;
      W_g[2,2] := -0.02538709;
      W_g[2,3] := -0.10518261;
      W_g[2,4] := -0.09690855;
      W_g[2,5] := 0.13110280;
      W_g[2,6] := 0.55399138;
      W_g[2,7] := -0.37729910;
      W_g[2,8] := -0.10455446;
      W_g[2,9] := -0.42354736;
      W_g[2,10] := 0.00632633;
      W_g[2,11] := 0.17120209;
      W_g[2,12] := -0.27252370;
      W_g[2,13] := -0.47738433;
      W_g[2,14] := -0.01380447;
      W_g[2,15] := -0.00504201;
      W_g[2,16] := 0.04669758;
      W_g[2,17] := -0.07789133;
      W_g[2,18] := -0.11861567;
      W_g[2,19] := -0.00203427;
      W_g[2,20] := 0.23830740;
      W_g[2,21] := 0.07300918;
      W_g[2,22] := 0.04740287;
      W_g[2,23] := -0.21146311;
      W_g[2,24] := -0.27551419;
      W_g[2,25] := -0.44383126;
      W_g[2,26] := -0.34758016;
      W_g[2,27] := 0.19908582;
      W_g[2,28] := 0.26224342;
      W_g[2,29] := -0.39878350;
      W_g[2,30] := 0.04991197;
      W_g[2,31] := 0.14302830;
      W_g[2,32] := -0.00475011;
      W_g[2,33] := -0.12771903;
      W_g[2,34] := -0.19415860;
      W_g[2,35] := 0.09121127;
      W_g[2,36] := -0.47490549;
      W_g[2,37] := 0.04646556;
      W_g[2,38] := -0.05770580;
      W_g[2,39] := -0.02702624;
      W_g[3,0] := 0.66790044;
      W_g[3,1] := -0.15152147;
      W_g[3,2] := -0.17599484;
      W_g[3,3] := 0.33776176;
      W_g[3,4] := -0.33888513;
      W_g[3,5] := 0.13354416;
      W_g[3,6] := -0.46012959;
      W_g[3,7] := 0.15908432;
      W_g[3,8] := -0.53887439;
      W_g[3,9] := -0.18714111;
      W_g[3,10] := -0.50302261;
      W_g[3,11] := -0.00954076;
      W_g[3,12] := 0.43053734;
      W_g[3,13] := 0.02114636;
      W_g[3,14] := 0.16980933;
      W_g[3,15] := -0.58761334;
      W_g[3,16] := 0.03133189;
      W_g[3,17] := -0.45295224;
      W_g[3,18] := 0.13907465;
      W_g[3,19] := 0.13671292;
      W_g[3,20] := 0.41902876;
      W_g[3,21] := 0.09891476;
      W_g[3,22] := -0.09855273;
      W_g[3,23] := 0.44152388;
      W_g[3,24] := -0.13008223;
      W_g[3,25] := -0.03226718;
      W_g[3,26] := -0.29500347;
      W_g[3,27] := -0.10089855;
      W_g[3,28] := 0.62393677;
      W_g[3,29] := 0.28965864;
      W_g[3,30] := -0.14991666;
      W_g[3,31] := 0.96139205;
      W_g[3,32] := 0.23747276;
      W_g[3,33] := 0.09901027;
      W_g[3,34] := 0.37833998;
      W_g[3,35] := -0.00466951;
      W_g[3,36] := 0.18169127;
      W_g[3,37] := 0.06343419;
      W_g[3,38] := -0.03238372;
      W_g[3,39] := 0.35362154;
      W_g[4,0] := -0.98030257;
      W_g[4,1] := 0.05196754;
      W_g[4,2] := 0.50153446;
      W_g[4,3] := 0.38619426;
      W_g[4,4] := 0.32922885;
      W_g[4,5] := -0.32188499;
      W_g[4,6] := 0.44783571;
      W_g[4,7] := -0.93163556;
      W_g[4,8] := 0.20751548;
      W_g[4,9] := -0.33809665;
      W_g[4,10] := 1.06782675;
      W_g[4,11] := -0.52386844;
      W_g[4,12] := 0.48961398;
      W_g[4,13] := -0.08319489;
      W_g[4,14] := 0.07775006;
      W_g[4,15] := 0.43782815;
      W_g[4,16] := -0.01010062;
      W_g[4,17] := -0.05047823;
      W_g[4,18] := 0.03664025;
      W_g[4,19] := -0.37702709;
      W_g[4,20] := 0.33760449;
      W_g[4,21] := 0.52333146;
      W_g[4,22] := 0.00913551;
      W_g[4,23] := 0.26169059;
      W_g[4,24] := 0.44963381;
      W_g[4,25] := 0.38881618;
      W_g[4,26] := -0.26409152;
      W_g[4,27] := -0.03092019;
      W_g[4,28] := -0.06874726;
      W_g[4,29] := 0.56894487;
      W_g[4,30] := 0.20915844;
      W_g[4,31] := 0.00012731;
      W_g[4,32] := 0.18578061;
      W_g[4,33] := 0.04220859;
      W_g[4,34] := 0.21296906;
      W_g[4,35] := 0.07501526;
      W_g[4,36] := 0.15391923;
      W_g[4,37] := 0.23479983;
      W_g[4,38] := 0.55838788;
      W_g[4,39] := 0.21783896;
      W_g[5,0] := 0.03072209;
      W_g[5,1] := 0.32084212;
      W_g[5,2] := 0.05682547;
      W_g[5,3] := -0.27383399;
      W_g[5,4] := -0.04110011;
      W_g[5,5] := -0.02305688;
      W_g[5,6] := 0.15270616;
      W_g[5,7] := -0.01929974;
      W_g[5,8] := -0.11035407;
      W_g[5,9] := 0.06503577;
      W_g[5,10] := 0.15678713;
      W_g[5,11] := 0.35518146;
      W_g[5,12] := -0.31208324;
      W_g[5,13] := -0.40173215;
      W_g[5,14] := -0.07717644;
      W_g[5,15] := -0.12580223;
      W_g[5,16] := 0.11613476;
      W_g[5,17] := -0.00657989;
      W_g[5,18] := 0.07340264;
      W_g[5,19] := -0.76857251;
      W_g[5,20] := -0.21624063;
      W_g[5,21] := 0.22518300;
      W_g[5,22] := 0.10625836;
      W_g[5,23] := 0.13706444;
      W_g[5,24] := -0.42099634;
      W_g[5,25] := -0.37740153;
      W_g[5,26] := 0.12714347;
      W_g[5,27] := -0.27696231;
      W_g[5,28] := -0.05975693;
      W_g[5,29] := -0.12939759;
      W_g[5,30] := 0.10944291;
      W_g[5,31] := 0.36755753;
      W_g[5,32] := -0.13962130;
      W_g[5,33] := -0.08474881;
      W_g[5,34] := -0.02089391;
      W_g[5,35] := -0.31487858;
      W_g[5,36] := 0.28444338;
      W_g[5,37] := -0.27468029;
      W_g[5,38] := 0.09558668;
      W_g[5,39] := -0.02762687;
      W_g[6,0] := 0.06528252;
      W_g[6,1] := -0.11730083;
      W_g[6,2] := 0.20279023;
      W_g[6,3] := 0.01967611;
      W_g[6,4] := 0.20667711;
      W_g[6,5] := -0.01244465;
      W_g[6,6] := -0.17045607;
      W_g[6,7] := 0.01241645;
      W_g[6,8] := -0.25576153;
      W_g[6,9] := -0.09515689;
      W_g[6,10] := 0.07613542;
      W_g[6,11] := 0.10648429;
      W_g[6,12] := -0.24497978;
      W_g[6,13] := -0.10179006;
      W_g[6,14] := 0.00171832;
      W_g[6,15] := -0.05910730;
      W_g[6,16] := 0.24741447;
      W_g[6,17] := -0.00957987;
      W_g[6,18] := 0.04504933;
      W_g[6,19] := 0.14365739;
      W_g[6,20] := 0.63776219;
      W_g[6,21] := -0.30890781;
      W_g[6,22] := -0.09165695;
      W_g[6,23] := 0.14273126;
      W_g[6,24] := -0.23289602;
      W_g[6,25] := -0.06301894;
      W_g[6,26] := -0.17733252;
      W_g[6,27] := -0.12566659;
      W_g[6,28] := -0.27798054;
      W_g[6,29] := 0.04181678;
      W_g[6,30] := -0.07146701;
      W_g[6,31] := -0.00828138;
      W_g[6,32] := -0.00004499;
      W_g[6,33] := -0.02710683;
      W_g[6,34] := -0.28370047;
      W_g[6,35] := 0.03627095;
      W_g[6,36] := 0.00073252;
      W_g[6,37] := 0.01647271;
      W_g[6,38] := -0.01837973;
      W_g[6,39] := -0.22433242;
      W_g[7,0] := 0.55378538;
      W_g[7,1] := 0.30619401;
      W_g[7,2] := 0.53044039;
      W_g[7,3] := 0.24350011;
      W_g[7,4] := 0.03852860;
      W_g[7,5] := -0.00226828;
      W_g[7,6] := -0.14655991;
      W_g[7,7] := -0.05021800;
      W_g[7,8] := 0.36482096;
      W_g[7,9] := -0.02399567;
      W_g[7,10] := -0.06456903;
      W_g[7,11] := 0.01613679;
      W_g[7,12] := -0.16384159;
      W_g[7,13] := -0.17693371;
      W_g[7,14] := 0.01647294;
      W_g[7,15] := 0.00100905;
      W_g[7,16] := -0.03387517;
      W_g[7,17] := -0.02685565;
      W_g[7,18] := -0.35300040;
      W_g[7,19] := 0.15475453;
      W_g[7,20] := 0.06111860;
      W_g[7,21] := 0.03696573;
      W_g[7,22] := 0.03331326;
      W_g[7,23] := 0.05765501;
      W_g[7,24] := 0.08704191;
      W_g[7,25] := 0.29588538;
      W_g[7,26] := 0.09131306;
      W_g[7,27] := -0.03710754;
      W_g[7,28] := 0.01770943;
      W_g[7,29] := -0.05923130;
      W_g[7,30] := 0.04210841;
      W_g[7,31] := 0.09924227;
      W_g[7,32] := -0.03344223;
      W_g[7,33] := -0.06622621;
      W_g[7,34] := 0.36641309;
      W_g[7,35] := -0.00420983;
      W_g[7,36] := -0.02636149;
      W_g[7,37] := -0.07082810;
      W_g[7,38] := -0.04731666;
      W_g[7,39] := 0.11440528;
      W_g[8,0] := -0.24883498;
      W_g[8,1] := 0.24131876;
      W_g[8,2] := 0.03446972;
      W_g[8,3] := -0.17805213;
      W_g[8,4] := -0.04451150;
      W_g[8,5] := 0.07381167;
      W_g[8,6] := 0.08678459;
      W_g[8,7] := 0.05011131;
      W_g[8,8] := 0.18668757;
      W_g[8,9] := 0.21342294;
      W_g[8,10] := -0.26045439;
      W_g[8,11] := 0.08760744;
      W_g[8,12] := 0.27040973;
      W_g[8,13] := 0.06985493;
      W_g[8,14] := 0.41351974;
      W_g[8,15] := -0.00667003;
      W_g[8,16] := 0.14276765;
      W_g[8,17] := 0.10061210;
      W_g[8,18] := -0.14089714;
      W_g[8,19] := -0.25550368;
      W_g[8,20] := 0.13017167;
      W_g[8,21] := -0.39635801;
      W_g[8,22] := -0.04880680;
      W_g[8,23] := -0.21499138;
      W_g[8,24] := 0.04412201;
      W_g[8,25] := 0.00883397;
      W_g[8,26] := -0.35899398;
      W_g[8,27] := 0.01892924;
      W_g[8,28] := -0.09143472;
      W_g[8,29] := -0.19829857;
      W_g[8,30] := -0.05133336;
      W_g[8,31] := 0.26230633;
      W_g[8,32] := 0.09470810;
      W_g[8,33] := 0.11210908;
      W_g[8,34] := 0.16554591;
      W_g[8,35] := 0.12200377;
      W_g[8,36] := 0.04580530;
      W_g[8,37] := 0.06629571;
      W_g[8,38] := -0.10643665;
      W_g[8,39] := 0.03629560;
      W_g[9,0] := -0.42790633;
      W_g[9,1] := 0.18710488;
      W_g[9,2] := 0.36177769;
      W_g[9,3] := 0.45072201;
      W_g[9,4] := -0.52714986;
      W_g[9,5] := 0.00028343;
      W_g[9,6] := -0.61539882;
      W_g[9,7] := 0.35529020;
      W_g[9,8] := -0.22070977;
      W_g[9,9] := 0.15130371;
      W_g[9,10] := 0.04521370;
      W_g[9,11] := 0.38444006;
      W_g[9,12] := -0.19535124;
      W_g[9,13] := -0.05019497;
      W_g[9,14] := -0.14246918;
      W_g[9,15] := -0.07645082;
      W_g[9,16] := 0.16795936;
      W_g[9,17] := 0.01235962;
      W_g[9,18] := 0.05418243;
      W_g[9,19] := -0.66316724;
      W_g[9,20] := -0.60060507;
      W_g[9,21] := -0.63958752;
      W_g[9,22] := -0.32650322;
      W_g[9,23] := 0.11281379;
      W_g[9,24] := -0.76775253;
      W_g[9,25] := -0.90051788;
      W_g[9,26] := -0.04093074;
      W_g[9,27] := 0.95141566;
      W_g[9,28] := 0.84178418;
      W_g[9,29] := 0.32648510;
      W_g[9,30] := -0.16123995;
      W_g[9,31] := -0.02454353;
      W_g[9,32] := 0.06485219;
      W_g[9,33] := 0.03735679;
      W_g[9,34] := -0.15660901;
      W_g[9,35] := 0.21646944;
      W_g[9,36] := -0.53633404;
      W_g[9,37] := 0.12129372;
      W_g[9,38] := -0.36001900;
      W_g[9,39] := 0.16128390;
      W_g[10,0] := 0.17666045;
      W_g[10,1] := -0.00918789;
      W_g[10,2] := -0.23106144;
      W_g[10,3] := -0.84316653;
      W_g[10,4] := -0.15785550;
      W_g[10,5] := 0.10649782;
      W_g[10,6] := -0.14947529;
      W_g[10,7] := 0.19670546;
      W_g[10,8] := 0.01153113;
      W_g[10,9] := 0.67161006;
      W_g[10,10] := -0.02482281;
      W_g[10,11] := -1.39040852;
      W_g[10,12] := 0.09316730;
      W_g[10,13] := -0.48327872;
      W_g[10,14] := 0.10523200;
      W_g[10,15] := -0.58414435;
      W_g[10,16] := 0.08219520;
      W_g[10,17] := 0.65659487;
      W_g[10,18] := -0.24748397;
      W_g[10,19] := 0.09048693;
      W_g[10,20] := 0.09783195;
      W_g[10,21] := 0.19360939;
      W_g[10,22] := -0.05255168;
      W_g[10,23] := 0.03202261;
      W_g[10,24] := -0.16167313;
      W_g[10,25] := 0.02797973;
      W_g[10,26] := -0.04574471;
      W_g[10,27] := -0.06924049;
      W_g[10,28] := 0.20432237;
      W_g[10,29] := 0.41537574;
      W_g[10,30] := -0.05165868;
      W_g[10,31] := -0.52141285;
      W_g[10,32] := 0.13948496;
      W_g[10,33] := 0.19479860;
      W_g[10,34] := -0.28982541;
      W_g[10,35] := 0.16944499;
      W_g[10,36] := 0.00522505;
      W_g[10,37] := 0.08370305;
      W_g[10,38] := -0.13435189;
      W_g[10,39] := -0.02312672;
      W_g[11,0] := 0.02013403;
      W_g[11,1] := 0.09134999;
      W_g[11,2] := 0.10191370;
      W_g[11,3] := -0.31639898;
      W_g[11,4] := 0.19775309;
      W_g[11,5] := -0.07690994;
      W_g[11,6] := 0.04381794;
      W_g[11,7] := -0.02134414;
      W_g[11,8] := -0.10884380;
      W_g[11,9] := 0.16108947;
      W_g[11,10] := 0.26612344;
      W_g[11,11] := 0.07906064;
      W_g[11,12] := -0.26956782;
      W_g[11,13] := 0.19898185;
      W_g[11,14] := -0.08008219;
      W_g[11,15] := 0.11739381;
      W_g[11,16] := -0.06613845;
      W_g[11,17] := 0.07276598;
      W_g[11,18] := -0.02100142;
      W_g[11,19] := 0.04329674;
      W_g[11,20] := -0.35718477;
      W_g[11,21] := -0.45652404;
      W_g[11,22] := 0.07382967;
      W_g[11,23] := -0.21277735;
      W_g[11,24] := 0.86212504;
      W_g[11,25] := 0.80017167;
      W_g[11,26] := 0.02575941;
      W_g[11,27] := 0.33303621;
      W_g[11,28] := -0.41469184;
      W_g[11,29] := -0.19018589;
      W_g[11,30] := -0.00447020;
      W_g[11,31] := 0.64252478;
      W_g[11,32] := 0.13424975;
      W_g[11,33] := 0.26267499;
      W_g[11,34] := 0.42238405;
      W_g[11,35] := 0.05826613;
      W_g[11,36] := -0.14534219;
      W_g[11,37] := 0.24092248;
      W_g[11,38] := 0.01456369;
      W_g[11,39] := -0.15360974;
      W_g[12,0] := -0.75018907;
      W_g[12,1] := 0.12156846;
      W_g[12,2] := -0.14797975;
      W_g[12,3] := 0.49666521;
      W_g[12,4] := 0.14742504;
      W_g[12,5] := -0.06025932;
      W_g[12,6] := -0.10514629;
      W_g[12,7] := 0.51666707;
      W_g[12,8] := -0.43515047;
      W_g[12,9] := 0.10338181;
      W_g[12,10] := 0.08973016;
      W_g[12,11] := -0.06708794;
      W_g[12,12] := -0.09652749;
      W_g[12,13] := -0.25314453;
      W_g[12,14] := 0.03715146;
      W_g[12,15] := -0.00260859;
      W_g[12,16] := -0.07890595;
      W_g[12,17] := -0.03232598;
      W_g[12,18] := -0.37715733;
      W_g[12,19] := 0.11189222;
      W_g[12,20] := 0.03655316;
      W_g[12,21] := 0.05601667;
      W_g[12,22] := 0.06752921;
      W_g[12,23] := 0.00744710;
      W_g[12,24] := 0.24519159;
      W_g[12,25] := 0.25994793;
      W_g[12,26] := 0.22617993;
      W_g[12,27] := -0.07020248;
      W_g[12,28] := -0.20237362;
      W_g[12,29] := -0.14392392;
      W_g[12,30] := 0.08102873;
      W_g[12,31] := -0.05696565;
      W_g[12,32] := 0.02835622;
      W_g[12,33] := -0.02322037;
      W_g[12,34] := 0.43416402;
      W_g[12,35] := -0.00790363;
      W_g[12,36] := -0.00377206;
      W_g[12,37] := -0.00598957;
      W_g[12,38] := -0.15154590;
      W_g[12,39] := 0.11662770;
      W_g[13,0] := -0.31849653;
      W_g[13,1] := 0.02676725;
      W_g[13,2] := 0.09364573;
      W_g[13,3] := -0.03316357;
      W_g[13,4] := -0.17901814;
      W_g[13,5] := 0.01395635;
      W_g[13,6] := -0.28069612;
      W_g[13,7] := 0.13494132;
      W_g[13,8] := 0.10521787;
      W_g[13,9] := 0.18218730;
      W_g[13,10] := -0.06014048;
      W_g[13,11] := 0.11842346;
      W_g[13,12] := -0.18528548;
      W_g[13,13] := 0.07218965;
      W_g[13,14] := -0.00519596;
      W_g[13,15] := -0.03343331;
      W_g[13,16] := 0.00436692;
      W_g[13,17] := 0.01997596;
      W_g[13,18] := -0.01004514;
      W_g[13,19] := 0.12576054;
      W_g[13,20] := 0.21994683;
      W_g[13,21] := 0.43556800;
      W_g[13,22] := -0.07989552;
      W_g[13,23] := 0.04946299;
      W_g[13,24] := -0.48828560;
      W_g[13,25] := -0.42732292;
      W_g[13,26] := -0.23599178;
      W_g[13,27] := 0.76446098;
      W_g[13,28] := -0.82037020;
      W_g[13,29] := 0.12914550;
      W_g[13,30] := -0.08376030;
      W_g[13,31] := 0.17175832;
      W_g[13,32] := -0.03239495;
      W_g[13,33] := -0.01117187;
      W_g[13,34] := -0.16287006;
      W_g[13,35] := -0.04970106;
      W_g[13,36] := 0.20778099;
